Omron Sysmac Studio project 04820KA001 Mono Slitter 903_V12_1105 (Sysmac Studio 1.60.0.64010, StandardProject)
(* Modified to Connect 2nd Diameter Sens *)

# Controller PLC: NX1P2-9024DT1 version 1.42
Units and slaves: Node1 : IL EC BK-PAC(E001); 0 : IB IL 24 DI 8/HD-ECO(M1); 1 : IB IL 24 DO 8/HD-ECO(M2); Unit 1 : NX-PF0730 (N3); Unit 2 : NX-AD2603 (N1); Unit 3 : NX-EC0122 (N2)
Task PrimaryTask (priority 4, period or condition 4000): TaglMonoTRM

VAR_GLOBAL
    Pot1_Work_Velocity : INT;  (* Potentiometer 1 value - Work speed -	Valore potenziometro 1 - Lavoro -; at BuiltInIO://opt/#0/Ch1_Analog_Input_Value; published *)
    InvRef : INT;  (* Inverter speed reference	Riferimento velocità inverter; at BuiltInIO://opt/#0/Ch2_Analog_Output_Value; published *)
    Fix10Vdc : INT;  (* Fixed 10 Vdc generator	Generatore 10Vdc fisso; at BuiltInIO://opt/#0/Ch1_Analog_Output_Value; published *)
END_VAR
VAR_GLOBAL RETAIN
    VelMax : REAL := 800;  (* Maximum speed	Velocità massima; published *)
END_VAR
VAR_GLOBAL
    VelSet : REAL;  (* Set speed	Velocità impostata; published *)
END_VAR
VAR_GLOBAL RETAIN
    RwSlowDecelK : REAL := 0.15;  (* Learned slow-down decel per mm of rewinder diameter (mm/s2 per mm); published *)
    RwMaxSlowFallback : REAL := 1285.0;  (* Rewinder max: slow-down diameter while K not learned (mm); published *)
END_VAR
VAR_GLOBAL
    PaperDensity : REAL;  (* published *)
END_VAR
VAR_GLOBAL RETAIN
    Language : DINT;  (* Language	Lingua; published *)
    RwThickMin_mm : REAL := 0.02;  (* Learning: min plausible paper thickness (mm); published *)
END_VAR
VAR_GLOBAL
    PulseRate : UDINT;  (* Pulses per 100 ms	Impulsi * 100ms; at IOBus://unit#3/Ch1 Pulse Rate; published *)
END_VAR
VAR_GLOBAL RETAIN
    RwThickMax_mm : REAL := 2.0;  (* Learning: max plausible paper thickness (mm); published *)
    RwDecelMin_mm : REAL := 20.0;  (* Learning: min plausible stop decel (mm/s2); published *)
    RwDecelMax_mm : REAL := 5000.0;  (* Learning: max plausible stop decel (mm/s2); published *)
    RwLearnFailMax : INT := 12;  (* Learning: failed windows before alarm (12 = 2 min); published *)
    RwStopFailMax : INT := 3;  (* Learning: failed stops before alarm; published *)
    RwThick_mm : REAL;  (* Learned paper thickness (mm); published *)
END_VAR
VAR_GLOBAL
    OverSpeed : BOOL;  (* Speed too high	Velocità troppo alta; published *)
END_VAR
VAR_GLOBAL RETAIN
    WorkSpd_Max : REAL := 500.0;  (* Work speed pot full scale (m/min), 50..VelMax; published *)
    WorkSpd_Max_Set : REAL := 400.0;  (* HMI request: work pot full scale (m/min), applied only with motor stopped; published *)
    UwRawMin : INT := 10;  (* Unwinder sonar raw min (below = sensor fault, alarm 17); published *)
    UwRawMax : INT := 3990;  (* Unwinder sonar raw max (above = sensor fault / no echo, alarm 17); published *)
    TensCheckEnable : BOOL := False;  (* Tension check ON (HMI switch); OFF = start as before; published *)
    TensWaitSpd : REAL := 10.0;  (* Speed held after START until tension established (m/min); published *)
END_VAR
VAR_GLOBAL
    TensionOK : BOOL := False;  (* Tension established (debounced T-one Alarm 0); published *)
    TensWait : BOOL := False;  (* Waiting for tension (speed held at TensWaitSpd, HMI lamp); published *)
    SonarAsk : BOOL := False;  (* V10 HMI popup: sonar is OFF, turn it on? (HMI NO resets it); published *)
END_VAR
VAR_GLOBAL RETAIN
    UwSlow_at_D_Req : BOOL := True;  (* V7c: unwinder diameter slow-down follows the speed (FALSE = fixed UwSlowDown_Diam); published *)
END_VAR
VAR_GLOBAL
    UwSlowDiamAct : REAL := 0.0;  (* V7c: unwinder slows down at this diameter (mm), HMI display; published *)
END_VAR
VAR_GLOBAL RETAIN
    FinalStopDecel : REAL := 500.0;  (* V12: end-of-roll stop ramp, web decel (mm/s2), 0 = drive DEC ramp as before, 50..2000; published *)
END_VAR
VAR_GLOBAL
    FinalStopRamp : BOOL := False;  (* V12: end-of-roll stop ramp running (HMI lamp); published *)
END_VAR
VAR_GLOBAL RETAIN
    RwJogMaxDiam : REAL := 400.0;  (* V7d: jog blocked above this rewinder diameter (mm), 0 = no limit; published *)
END_VAR
VAR_GLOBAL
    JogInhibit : BOOL := False;  (* V7d: jog blocked (rewinder roll too big), HMI lamp; published *)
END_VAR
VAR_GLOBAL RETAIN
    SCurveTime : REAL := 0.5;  (* V7f: S-curve rounding of the AUTO ramps (s), 0 = off, max 2; published *)
END_VAR
VAR_GLOBAL
    TOneDecel : BOOL := False;  (* V7f: line decelerating (for a T-one stop/boost input); published *)
END_VAR
VAR_GLOBAL RETAIN
    HornStartBeep_s : REAL := 1.0;  (* V9 horn: beep when the slow-down starts (s), 0 = off, max 5; published *)
    HornBeepLen_s : REAL := 0.2;  (* V9 horn: length of the short beeps during slow-down (s), 0 = off, max 2; published *)
    HornBeepPeriod : REAL := 5.0;  (* V9 horn: one short beep every ... s during slow-down, 0 = off, max 30; published *)
    HornStopBeep_s : REAL := 3.0;  (* V9 horn: beep when stopped after a slow-down (s), 0 = off, max 10; published *)
END_VAR
VAR_GLOBAL
    HornTest : BOOL := False;  (* V9 horn: HMI test button (momentary), machine stopped only; published *)
END_VAR
VAR_GLOBAL RETAIN
    RwLockDiam : REAL := 300.0;  (* V9: paper thickness LOCKED at this rewinder diameter (mm), 0 = never lock; published *)
    RwLockMinGrow_mm : REAL := 50.0;  (* V9: min diameter growth since the start of learning before locking (mm); published *)
    RwMatLocked : BOOL := False;  (* V9: paper thickness locked (HMI lamp), NEW PAPER / GSM YES unlocks; published *)
END_VAR
VAR_GLOBAL
    LongThick_mm : REAL := 0.0;  (* V9: thickness from the long baseline (mm), HMI display; published *)
    RwDiamRev : REAL := 0.0;  (* V9: rewinder diameter averaged over one revolution (mm); published *)
    RwWave_mm : REAL := 0.0;  (* V9: diameter wave peak-peak in the last revolution (mm), HMI; published *)
    UwStopLenShow : BOOL := False;  (* V9 HMI: show unwinder STOP LENGTH (AUTO STOP UNWINDER active); published *)
    UwSlowDiamShow : BOOL := False;  (* V9 HMI: show unwinder SLOW AT diameter (normal operation, sonar ON); published *)
END_VAR
VAR_GLOBAL RETAIN
    SoftCancelAccel : REAL := 100.0;  (* V9: then ramp up at this web accel (mm/s2), 0 = AccelWeb; published *)
END_VAR
VAR_GLOBAL
    RwMatReset : BOOL := False;  (* HMI NEW PAPER: forget the learned paper thickness RwMat_K (PLC resets it); published *)
END_VAR
VAR_GLOBAL RETAIN
    FinalSpd_Max_Set : REAL := 80.0;  (* HMI request: final pot full scale (m/min), applied only with motor stopped; published *)
    FinalSpd_Max : REAL := 80.0;  (* Final speed pot full scale (m/min), 5..WorkSpd_Max; published *)
END_VAR
VAR_GLOBAL
    UnderSpeed : BOOL;  (* Speed too low	Velocità troppo bassa; published *)
    RwLearnReset : BOOL := False;  (* HMI / Watch: clear learned decels RwStopDecelK, RwStopDecel, RwSlowDecelK (PLC resets it); published *)
END_VAR
VAR_GLOBAL RETAIN
    RwCoreDiameter : REAL := 100.0;  (* Rewinder core outside diameter for TEACH CORE (mm); published *)
END_VAR
VAR_GLOBAL
    RwTeachCore : BOOL := False;  (* HMI: TEACH CORE request (PLC resets it); published *)
    RwTeachState : INT := 0;  (* TEACH CORE: 0 idle 1 teaching 2 done 3 refused; published *)
END_VAR
VAR_GLOBAL RETAIN
    SpdDelta_Percent : REAL := 12.0;  (* Speed difference percentage	Percentuale differenza velocità; published *)
END_VAR
VAR_GLOBAL
    Encoder_Pos : DINT;  (* Encoder counter	Contatore encoder; at IOBus://unit#3/Ch1 Encoder Present Position; published *)
    UwTeachState : INT := 0;  (* Unwinder TEACH CORE: 0 idle 1 teaching 2 done 3 refused; published *)
    Encoder_On : BOOL;  (* Encoder enable	Abilita encoder; at IOBus://unit#3/Ch1 Encoder Counter Operation Command/Ch1 Counter Enable; published *)
    Encoder_Reset : BOOL;  (* Encoder reset	Reset encoder; at IOBus://unit#3/Ch1 Encoder Counter Operation Command/Ch1 Internal Reset Execution; published *)
    HMI_Screen : ARRAY[0..1] OF DINT;  (* HMI panel Screen	Pagina pannello; published *)
END_VAR
VAR_GLOBAL RETAIN
    Velocity_M_min : REAL;  (* Speed in m/min	Velocità in mt/min; published *)
    Current_Metre : REAL;  (* Current metres	Metri attuali; published *)
END_VAR
VAR_GLOBAL
    I_RsetCnt : BOOL;  (* Metre counter reset button	Pulsante reset contametri; published *)
END_VAR
VAR_GLOBAL RETAIN
    Speed_Display : REAL;  (* Set speed (displayed)	Velocità impostata visualizzata; published *)
END_VAR
VAR_GLOBAL
    I_ControlVoltage : BOOL;  (* In_0 ControlVoltageON	Ausiliari inseriti; at BuiltInIO://cpu/#0/Input_Bit_00; published *)
    I_Start_PB : BOOL;  (* In_1 Start button	Pulsante di marcia; at BuiltInIO://cpu/#0/Input_Bit_01; published *)
    I_Stop_PB : BOOL;  (* In_2 Stop button	Pulsante di arresto; at BuiltInIO://cpu/#0/Input_Bit_02; published *)
    I_Motor_Thermal : BOOL;  (* In_3 Motor thermal switch	Pastiglia termica motore; at BuiltInIO://cpu/#0/Input_Bit_03; published *)
    I_Prot_ByPass : BOOL;  (* In_4 Guards-bypassed selector switch - Under Panel	Selettore protezioni escluse; at BuiltInIO://cpu/#0/Input_Bit_04; published *)
    I_Hub_Position : BOOL;  (* In_5 Hub/chuck in extraction position	Mozzo in posizione di estrazione; at BuiltInIO://cpu/#0/Input_Bit_05; published *)
    I_FrontGuard_Closed : BOOL;  (* In_6 Front guard closed	Riparo frontale chiuso; at BuiltInIO://cpu/#0/Input_Bit_06; published *)
    I_Jog_PB : BOOL;  (* In_7 Jog Push button	Pulsante velocità ridotta; at BuiltInIO://cpu/#0/Input_Bit_07; published *)
    I_VFD_Alarm : BOOL;  (* In_8 Inverter in alarm	Inverter in allarme; at BuiltInIO://cpu/#0/Input_Bit_08; published *)
    I_Side_Door_Closed : BOOL;  (* In_Side Door is Closed	Fotocellula diametro bobina; at BuiltInIO://cpu/#0/Input_Bit_13; published *)
    I_OR_Position_Sens : BOOL;  (* OverRider position sens	Sensore posizione pressore; at ECAT://node#[1,0]/IB IL 24 DI 8/HD-ECO Input-_IN01 (Pin 1.1)_6000_01; published *)
    I_OR_Hoover_Mode : BOOL;  (* OverRider Hoover Mode	Pressostato pressore; at ECAT://node#[1,0]/IB IL 24 DI 8/HD-ECO Input-_IN02 (Pin 2.1)_6000_02; published *)
    I_OR_Auto_OS : BOOL;  (* OverRider in automatic	Pressore in automatico; at ECAT://node#[1,0]/IB IL 24 DI 8/HD-ECO Input-_IN03 (Pin 1.2)_6000_03; published *)
    I_OR_Cont_OS : BOOL;  (* OverRider in continuous	Pressore in continuo; at ECAT://node#[1,0]/IB IL 24 DI 8/HD-ECO Input-_IN04 (Pin 2.2)_6000_04; published *)
    O_MotorStart : BOOL;  (* Q_0 Motor start	Start motore; at BuiltInIO://cpu/#0/Output_Bit_00; published *)
    I_FanTemp_Ok : BOOL;  (* Motor (fan) thermal OK	Termico motore ok; at ECAT://node#[1,0]/IB IL 24 DI 8/HD-ECO Input-_IN06 (Pin 2.3)_6000_06; published *)
    O_Alarm_Array : BOOL;  (* Alarm lamp	Lampada allarme; at ECAT://node#[1,1]/IB IL 24 DO 8/HD-ECO Output_OUT01 (Pin 1.1)_7000_01; published *)
    O_Prot_ByPass_Lamp : BOOL;  (* Guards bypassed lamp	Lampada protezioni escluse; published *)
    O_Motor_Lamp : BOOL;  (* Q_1 Motor ON lamp	Lampada motore on; at BuiltInIO://cpu/#0/Output_Bit_01; published *)
    O_RwUnload : BOOL;  (* Unloaders enable - opening	Consenso a scaricatori in apertura; at ECAT://node#[1,1]/IB IL 24 DO 8/HD-ECO Output_OUT03 (Pin 1.2)_7000_03; published *)
    O_FrontGuard_ByPass : BOOL;  (* Front guard bypass	Bypass protezione frontale; at ECAT://node#[1,1]/IB IL 24 DO 8/HD-ECO Output_OUT04 (Pin 2.2)_7000_04; published *)
    O_Brake : BOOL;  (* Q_2 Brake command	Comando freno; at BuiltInIO://cpu/#0/Output_Bit_02; published *)
    O_OR_Auto_Lamp : BOOL;  (* Q_6 OverRider auto/continuous lamp	Lamapda pressore in auto o continuo; at BuiltInIO://cpu/#0/Output_Bit_06; published *)
    O_OverRider_Up : BOOL;  (* Q_9 Raise OverRider ~10mm Over Rewinder roll	Solleva pressore; at BuiltInIO://cpu/#0/Output_Bit_09; published *)
    O_OverRider_Hold : BOOL;  (* Q_4 OverRider Lock 	Blocca pressore; at BuiltInIO://cpu/#0/Output_Bit_04; published *)
    O_CoolingFan : BOOL;  (* Q_3 Brake and motor fans	Ventole freno e motore; at BuiltInIO://cpu/#0/Output_Bit_03; published *)
END_VAR
VAR_GLOBAL RETAIN
    Fan_Timeout : REAL := 0.5;  (* Fans stop timeout [min]	Timeout stop ventole da pannello; published *)
    OverRider_TimeOFF : REAL := 0.01;  (* OverRider photocell OFF timeout (panel)	Timeout fotocellula pressore off; published *)
    OverRider_TimeON : REAL := 0.05;  (* OverRider photocell ON timeout (panel)	Timeout fotocellula pressore on; published *)
END_VAR
VAR_GLOBAL
    AlarmOn : BOOL;  (* Alarm active	Allarme presente; published *)
    BuzzerOn : BOOL;  (* Panel buzzer command	Comando buzzer pannello; published *)
    Msg : INT;  (* Message	Messagio; published *)
    Index_B : INT;  (* Alarm index	Indice allarme; published *)
    MotStop : BOOL;  (* Motor stopped	Motore fermo; published *)
    Clock1s : BOOL;  (* 1 s clock	Clock di 1s; published *)
END_VAR
VAR_GLOBAL RETAIN
    ManMode : BOOL;  (* Manual mode	Modo manuale; published *)
END_VAR
VAR_GLOBAL
    Counter_Reset : BOOL;  (* Counter reset from panel	Reset contatore da pannello; published *)
    I_FrontGuard_Open : BOOL;  (* In_9 Front guard open	Riparo frontale aperto; at BuiltInIO://cpu/#0/Input_Bit_09; published *)
    O_RwLoading_Enable : BOOL;  (* Q_7 Unloaders Load enable - closing	Consenso scaricatori in chiusura; at BuiltInIO://cpu/#0/Output_Bit_07; published *)
END_VAR
VAR_GLOBAL RETAIN
    JogSpd_SP : REAL := 10.0;  (* Speed in manual	Velocità in manuale; published *)
END_VAR
VAR_GLOBAL
    O_AccDec2 : BOOL;  (* Q_5 Second acc/dec ramp	Seconda rampa di acc/dec; at BuiltInIO://cpu/#0/Output_Bit_05; published *)
END_VAR
VAR_GLOBAL RETAIN
    AccelTrim : REAL := 0.08;  (* Acceleration coefficient in run	Coefficente accelerazione in lavoro; published *)
    DecelTrim : REAL := 0.08;  (* Deceleration coefficient in run	Coefficente decelerazione in lavoro; published *)
    DecelCoarse : REAL := 0.3;  (* Acceleration coefficient at start (orig. comment; name suggests decel)	Coefficente accelerazione in partenza; published *)
    AccelCoarse : REAL := 0.3;  (* Acceleration coefficient at start (orig. comment; name suggests accel)	Coefficente decelerazione in partenza; published *)
END_VAR
VAR_GLOBAL
    UwStopDiamShow : BOOL := False;  (* V11 HMI: show unwinder STOP AT diameter (slow-down reached, decel / final speed); published *)
    O_AcousticSignal : BOOL;  (* Q_8 Horn / Acoustic signal	Segnalatore acustico; at BuiltInIO://cpu/#0/Output_Bit_08; published *)
    Pot2_Slow_Velocity : INT;  (* Potentiometer 2 value - Final speed -	Valore potenziometro 2 - Finale -; at BuiltInIO://opt/#0/Ch2_Analog_Input_Value; published *)
    I_AutoStop_OS : BOOL;  (* In_10 Stop on metre counter	Arresto con contametri; at BuiltInIO://cpu/#0/Input_Bit_10; published *)
    I_Input_11_Spare_1255 : BOOL;  (* In_11 SPARE  (wire 12.55) Under Panel	Rallento a fine bobina; at BuiltInIO://cpu/#0/Input_Bit_11 *)
    I_WebBreak_Monitor : BOOL;  (* In_12 Paper break monitoring ON	Controllo rottura carta on; at BuiltInIO://cpu/#0/Input_Bit_12; published *)
    I_Vacuum_OK : BOOL;  (* Extractor fan thermal OK	Termico aspiratore ok; at IOBus://unit#3/Ch1 Reset/External Input Status/Ch1 External Input 0 Status; published *)
    I_T_one_TensionOK : BOOL;  (* T-one Alarm 0 (15-16): tension established (replaces I_SlowSens_PH); at ECAT://node#[1,0]/IB IL 24 DI 8/HD-ECO Input-_IN05 (Pin 1.3)_6000_05; published *)
    I_WebBreak_PH : BOOL;  (* Paper break photocell	Fotocellula rottura carta; at ECAT://node#[1,0]/IB IL 24 DI 8/HD-ECO Input-_IN07 (Pin 1.4)_6000_07; published *)
END_VAR
VAR_GLOBAL RETAIN
    UwStop_at_M_Val : REAL := 5100;  (* Unwinder Stop at metres	Metri totali; published *)
    UwSlowMargin_m : REAL := 10;  (* Unwinder Slow-down metres	Metri rallentamento; published *)
    LowSpd_Display : REAL;  (* Slow-down speed (displayed)	Velocità rallentamento visualizzata; published *)
    RwMaxDiam : REAL := 1315.0;  (* Rewinder max diameter protection (mm); published *)
END_VAR
VAR_GLOBAL
    RwMaxStop : BOOL;  (* Rewinder max diameter STOP (latched); published *)
END_VAR
VAR_GLOBAL RETAIN
    Encoder_Pulse : INT := 1000;  (* Encoder pulses/Rotation	Impulsi encoder; published *)
    RwSlowDecelLrn : REAL := 0.0;  (* Learned real slow-down decel (mm/s2) - 0 = not learned; published *)
END_VAR
VAR_GLOBAL
    CountReset_Req : BOOL;  (* Counter reset requested	Richiesto reset contatore; published *)
    Psw : INT;  (* Password Entry	Password; published *)
    I_RsetAlarm : BOOL;  (* Alarm reset	Reset allarmi; at ECAT://node#[1,0]/IB IL 24 DI 8/HD-ECO Input-_IN08 (Pin 2.4)_6000_08; published *)
END_VAR
VAR_GLOBAL RETAIN
    EncoderWheel_Circumf : REAL := 402;  (* Encoder wheel (Cylinder / Roller) Circumference [mm]	Diametro ruota encoder; published *)
END_VAR
VAR_GLOBAL
    AlarmCodeSV : ARRAY[0..32] OF BOOL;  (* Panel alarms	Allarmi a pannello; published *)
    SafeGuard_ByPass : BOOL;  (* Guards bypassed	Protezioni escluse; published *)
    FrontGuard_Closed : BOOL;  (* Front guard closed	Riparo frontale chiuso; published *)
    SoftStop : BOOL := False;  (* Soft stop in progress (HMI); published *)
END_VAR
VAR_GLOBAL RETAIN
    SoftStopEnable : BOOL := True;  (* STOP button = soft stop (False = immediate as before); published *)
    SoftStopEndSpd : REAL := 8.0;  (* Soft stop: run command drops below this speed (m/min); published *)
    UwDiam_Measure : REAL;  (* Measured distance	Distanza letta; published *)
    UwCoreDiameter : REAL := 100;  (* Core Outside diameter [mm]; published *)
    Core_Measure : BOOL := False;  (* Stored core value; published *)
    UwCoreDistance : REAL := 785.56;  (* Sonar distance to empty core. [mm]; published *)
END_VAR
VAR_GLOBAL
    AI_Diam_Unwinder : INT;  (* Analog value - UnWinder Diameter	Valore analogico misura bobina madre; at IOBus://unit#2/Ch1 Analog Input Value; published *)
END_VAR
VAR_GLOBAL RETAIN
    Measure_ON : BOOL := True;  (* Measurement enabled; published *)
    UwDiam_Act : REAL;  (* Measured roll diameter; published *)
    UwSlow_at_D_Val : REAL := 200;  (* Unwinder Slow-down diameter [mm]; published *)
    UwStopDiam_Limit : REAL := 110;  (* Stop diameter; published *)
END_VAR
VAR_GLOBAL
    Alarm_Reset : BOOL;  (* Alarm reset from panel; published *)
    Psw22 : BOOL;  (* Password 22 for Popup 22; published *)
    Psw44 : BOOL;  (* Password 44 for Popup 44; published *)
    I_Roll_OK : BOOL;  (* Roll OK / Broken Holder Joint; published *)
    AI_Diam_Rewinder : INT;  (* Analog value - ReWinder Diameter; at IOBus://unit#2/Ch2 Analog Input Value; published *)
END_VAR
VAR_GLOBAL RETAIN
    RwStopEnable : BOOL := False;  (* Rewinder diameter stop enabled; published *)
    RwTargetDiam : REAL := 300.0;  (* Rewinder final diameter (mm); published *)
    RwUseSlow : BOOL := True;  (* Slow down before target; published *)
    RwSlowMargin_m : REAL := 10.0;  (* Rewinder Metres at slow speed before stop; published *)
    RwSlowDecel : REAL := 0.0;  (* Rewinder Slow-down decel mm/s2 - 0 = auto from DecStart; published *)
    RwResetHyst : REAL := 50.0;  (* Reset requests below target - this [mm]; published *)
    RwDist0V : REAL := 0.0;  (* DT35 distance at 0 V (mm); published *)
    RwDist10V : REAL := 782.0;  (* DT35 distance at 10 V (mm); published *)
    RwRawMin : INT := 10;  (* Raw below = sensor fault; published *)
    RwRawMax : INT := 3900;  (* Raw above = sensor fault; published *)
END_VAR
VAR_GLOBAL
    RwStopOnFault : BOOL := True;  (* Stop on sensor fault; published *)
END_VAR
VAR_GLOBAL RETAIN
    RwAxisDist : REAL := 727.0;  (* Sensor to shaft centre (mm) - teach; published *)
    RwFilter_K : REAL := 0.2;  (* Distance filter per 100 ms (0..1); published *)
    RwMinPulses : DINT := 1000;  (* Min pulses in window to learn; published *)
    RwLearn_K : REAL := 0.3;  (* Material factor filter weight; published *)
    RwMat_K : REAL := 0.0;  (* Learned material factor; published *)
    RwLearnStop : BOOL := True;  (* Learn stop decel on every stop; published *)
    RwMinLearnSpd : REAL := 15.0;  (* Min speed to learn a stop (m/min); published *)
    RwStopDecel : REAL := 0.0;  (* Learned stop decel (pulses/s2); published *)
    RwTreact : REAL := 0.03;  (* Stop reaction time (s); published *)
    RwTstopDef : REAL := 3.0;  (* Stop time until decel learned (s); published *)
    RwTrim : REAL := 1.0;  (* Stop length trim (>1 = earlier); published *)
END_VAR
VAR_GLOBAL
    RwDist : REAL;  (* Filtered distance (mm); published *)
    RwDiam : REAL;  (* Rewinder diameter (mm); published *)
    RwSpeed : REAL;  (* Line speed from encoder (m/min); published *)
    RwRemain_m : REAL;  (* Metres to target diameter; published *)
    RwStopLen_m : REAL;  (* Stopping length now (m); published *)
    RwSlowLen_m : REAL;  (* Rewinder Slow-down length [m]; published *)
    RwStop_at_D_Req : BOOL;  (* Rewinder diameter STOP request; published *)
    RwSlow_at_D_Req : BOOL;  (* Rewinder diameter SLOW request; published *)
    RwSensFault : BOOL;  (* Rewinder DT35 sensor fault; published *)
END_VAR
VAR_GLOBAL RETAIN
    UwStopEnable : BOOL := False;  (* Unwinder Auto Stop - Enable; published *)
END_VAR
VAR_GLOBAL
    SlowAtDisp : REAL;  (* HMI: slow-down starts at (m or mm, see SlowAtMode); published *)
    SlowAtMode : INT;  (* HMI: 0=none 1=unwinder [m] 2=rewinder [mm]; published *)
    SlowAtShow : BOOL;  (* HMI: show slow-down display; published *)
    UwSlow_at_M_Val : REAL;  (* Unwinder: slow-down starts at [m]; published *)
    UwSlow_at_M_Req : BOOL;  (* Unwinder metre slow-down request (latched); published *)
    RwSlow_at_D_Val : REAL;  (* Rewinder slow-down starts at diameter [mm]; published *)
    RwStop_at_D_Val : REAL;  (* Rewinder: stop command at diameter (mm); published *)
    RwMaxSlow : BOOL;  (* Rewinder max diameter SLOW (latched); published *)
END_VAR
VAR_GLOBAL RETAIN
    UwEmptyHyst : REAL := 30.0;  (* Unwinder Empty Hysteresis; published *)
END_VAR
VAR_GLOBAL
    GSM_Learned_OK : BOOL;  (* Paper [Grams / Square Meter]  FALSE until GSM learned; published *)
    RwMaxSlowAtDiam : REAL := 1370.0;  (* Rewinder max: slow-down starts at diameter (mm); published *)
END_VAR
VAR_GLOBAL RETAIN
    RwStopDecelK : REAL := 0.0;  (* Learned stop decel per mm of rewinder diameter (mm/s2 per mm); published *)
    SoftStopDecel : REAL := 500.0;  (* Soft stop decel (mm/s2), 0 = DecelCoarse; published *)
END_VAR
VAR_GLOBAL
    SpdMax_Pending : BOOL := False;  (* New pot range waiting for the motor to stop; published *)
END_VAR
VAR_GLOBAL RETAIN
    RwAxisDist_Prev : REAL := 727.0;  (* Rewinder: RwAxisDist before the last TEACH (for UNDO); published *)
    UwCoreDist_Prev : REAL := 785.56;  (* Unwinder: UwCoreDistance before the last TEACH (for UNDO); published *)
END_VAR
VAR_GLOBAL
    RwTeachUndo : BOOL := False;  (* HMI: UNDO rewinder TEACH (PLC resets it); published *)
    UwTeachUndo : BOOL := False;  (* HMI: UNDO unwinder TEACH (PLC resets it); published *)
    Psw33 : BOOL;  (* Password 33 for Popup 33; published *)
END_VAR
VAR_GLOBAL RETAIN
    RwMatChangePct : REAL := 35.0;  (* Paper change detection: window deviation (%), 2 windows in a row = new paper, 0 = off; published *)
    RwSlowFallbackMm : REAL := 30.0;  (* Rewinder: slow-down this many mm before the target while the paper thickness is not learned (0 = off); published *)
    RwAutoMaxSpd : REAL := 500.0;  (* Rewinder AUTO stop ON: maximum work speed (m/min), 0 = no limit; published *)
    RwWinLen_m : REAL := 60.0;  (* Paper thickness learning: MAX window length (m of paper); published *)
    RwWinGrow_mm : REAL := 5;  (* Paper thickness learning: window = this diameter growth (mm), 4 m .. RwWinLen_m; published *)
END_VAR
VAR_GLOBAL
    GsmAsk : BOOL := False;  (* HMI popup: new parent roll, did you change the paper? (HMI NO resets it); published *)
    GsmAskYes : BOOL := False;  (* HMI popup YES: forget the learned thickness (PLC resets it); published *)
END_VAR
VAR_GLOBAL RETAIN
    DecelWeb : REAL := 250.0;  (* V7: AUTO decel ramp, real web mm/s2 (0 = DecelCoarse); published *)
    AccelWeb : REAL := 200.0;  (* AUTO accel ramp, real web mm/s2 (0 = AccelCoarse); published *)
    RwRatioD : REAL := 3366.0;  (* V7: drive counts per m/min x rewinder diameter (mm), adapted while running; published *)
    FFEnable : BOOL := True;  (* V7: feed-forward speed loop ON (FALSE = old loop of rung 16); published *)
END_VAR
VAR_GLOBAL
    SpdHold : BOOL := False;  (* V9: speed held after START during a soft stop, START again = ramp up (HMI lamp); published *)
    SonarAskYes : BOOL := False;  (* V10 HMI popup YES: sonar ON (PLC resets it); published *)
    UwStop_at_D_Val : REAL := 0.0;  (* V11: unwinder stop command diameter (mm) so the web stops at UwDiamStop, HMI "STOP AT"; published *)
    Clock10ms : BOOL;  (* 10mS clock; published *)
    Clock100ms : bool;  (* 100mS clock; published *)
    Sec_to_Min : REAL;
    Psw48 : BOOL;  (* Password 48 for Popup 48; published *)
    JogRun : BOOL;  (* V10: JOG really running (button, not a normal run, not a soft stop); published *)
    GuardStopOK : BOOL;  (* V11: stopped for real -> guard bypass allowed (Output 13); published *)
    SlowDown : BOOL;  (* Slow down	Rallenta; published *)
    WarningOn : bool;  (* HMI Warning Display; published *)
    AlarmSilenced : BOOL;  (* published *)
END_VAR
VAR_GLOBAL RETAIN
    PaperGSM : REAL;  (* published *)
    WebWidth_mm : REAL;  (* published *)
    TensFactor : REAL;  (* Tension Helper; published *)
    TensShowKg : BOOL;  (* Tension Helper; published *)
    TensShowLb : BOOL;  (* Tension Helper; published *)
    TensShowN : BOOL;  (* Tension Helper; published *)
    TensIdeal_Disp : REAL;  (* Tension Helper; published *)
    TensUnit : INT;  (* Tension Helper; published *)
END_VAR
VAR_GLOBAL
    TensUnitPB : BOOL;  (* Tension Helper; published *)
    TensLostWarn : BOOL := False;  (* Tension lost while running (warning); published *)
    UwSensTest : BOOL := False;  (* Unwinder sonar fault (raw out of range 1 s); published *)
    UwSensFault : BOOL;  (* UnWinder Sensor Fault; published *)
    Thickness_Fault : BOOL;  (* Thickness Not Learned !; published *)
    AutoStopWhy : INT;  (* published *)
    AutoStopDone : BOOL;  (* published *)
    AutoEnRefused : BOOL;  (* published *)
    AutoEnWhy : INT;  (* published *)
END_VAR

PROGRAM TaglMonoTRM
VAR
    SpdDelta : REAL;  (* Minimum or maximum speed SpdDeltaerence	Minima o massima differenza velocità *)
    UwSlowDiamCalc : REAL;  (* V7c: speed-dependent unwinder slow-down diameter (mm) *)
    SonarRunMem : bool;
    EndStopReq : BOOL;  (* V12: end-of-roll stop requested (AutoStopCmd or unwinder diameter) *)
    Buffer_R : BOOL;  (* Buffer Result *)
    EndRampOK : BOOL;  (* V12: end-of-roll ramp usable (FinalStopDecel, FF active, running) *)
    EndRampHard : BOOL;  (* V12: safety net during the ramp -> immediate stop *)
    EndStopNow : BOOL;  (* V12: immediate end-of-roll stop (Motor_Manager rung 4) *)
    SonarInit : bool;
    UwSlowDiamLatch : BOOL;  (* V7c: unwinder diameter slow-down reached (frozen) *)
    FFRate : REAL;  (* V7f: ramp rate (reference per 4 ms scan) *)
    FFRateSet : REAL;  (* V7f: rate allowed to still stop at the target *)
    FFJerk : REAL;  (* V7f: max rate change per scan *)
    SpdScanCnt : INT;  (* V9: scan counter for the 100 ms speed window *)
    HornRun : BOOL;  (* V9: slow-down / final speed running *)
    HornRunMem : BOOL;  (* V9: edge memory *)
    HornStartMem : BOOL;  (* V9: start edge memory *)
    HornTicks : INT;  (* V9: scans since slow-down start *)
    HornCnt : INT;  (* V9: scans in the beep period *)
    HornPer : INT;  (* V9: beep period in scans *)
    HornStartScans : INT;  (* V9: start beep in scans *)
    HornLenScans : INT;  (* V9: short beep in scans *)
    HornSlowBeep : BOOL;  (* V9: slow-down beep *)
    HornStopPend : BOOL;  (* V9: stopped after a slow-down, waiting for standstill *)
    HornStopTicks : INT;  (* V9: stop beep counter *)
    LongActive : BOOL;  (* V9: long-baseline learning running *)
    LongValid : BOOL;  (* V9: long baseline >= 20 mm growth, replaces the windows *)
    LongStartPos : DINT;  (* V9: encoder at the start of the long baseline *)
    LongStartD : REAL;  (* V9: rewinder diameter at the start (mm) *)
    LongGrow_mm : REAL;  (* V9: growth since the start (mm) *)
    LongPls : REAL;  (* V9: pulses since the start *)
    LongK : REAL;  (* V9: K from the long baseline *)
    RevW : REAL;  (* V9: encoder pulses summed in the current revolution *)
    RevDP : DINT;  (* V9: encoder pulses this scan *)
    RevPrevPos : DINT;  (* V9: encoder last scan *)
    RevSum : REAL;  (* V9: sum of raw DT35 distance x pulses *)
    RevMin : REAL;  (* V9: min raw distance in the revolution *)
    RevMax : REAL;  (* V9: max raw distance in the revolution *)
    RwDiamRevOk : BOOL;  (* V9: one full revolution averaged since the last fault *)
    UwEmptyTicks : INT;  (* V9: unwinder empty time (100 ms ticks) *)
    UwFullTicks : INT;  (* V9: new roll seen time (100 ms ticks) *)
    GsmArmed : BOOL;  (* V9: roll was empty -> next new roll asks the GSM question *)
    T_JogStartBlk : TOF;  (* V9: START blocked while JOG held + 2 s *)
    StartHeldBlk : BOOL;  (* V9: START pressed during the block, wait for release *)
    StartPB_OK : BOOL;  (* V9: START push-button accepted (replaces I_Start_PB in General 7/8/10) *)
    FFSoftMem : BOOL;  (* V9: soft stop last scan (rung B) *)
    FFSlowAcc : BOOL;  (* V9: gentle ramp-up after a cancelled soft stop *)
    FFStartEdge : BOOL;  (* V9: START push-button edge (rung B) *)
    FFStartMem : BOOL;  (* V9: START last scan (rung B) *)
    SpdDeltaMin : REAL;  (* Minimum speed difference	Minima differenza velocità *)
    FFSqrtArg : REAL;  (* SQRT argument (REAL) *)
    SpdDeltaMax : REAL;  (* Maximum speed SpdDeltaerence	Massima differenza velocità *)
    SoftStopMem : BOOL;  (* v6r: soft stop edge memory *)
    SoftStopRatio : REAL;  (* v6r: InvRef counts per m/min, frozen at the soft stop start *)
    MemPos : DINT;  (* Previous encoder count	Contatore encoder precedente *)
    MatChangeCnt : INT;  (* v6s: consecutive learning windows far from RwMat_K *)
    DeltaPulse : DINT;  (* Encoder count difference	Differenza contatore encoder *)
    SlowMem : BOOL;  (* SlowDown edge memory *)
    DecelDiam : REAL;  (* Rewinder diameter used by the decel model (mm, min 100) *)
    TeachSwap : REAL;  (* Temporary for UNDO swap *)
    SlowStartDiam : REAL;  (* Diameter at slow-down start (mm) *)
    BrakeHold : BOOL;  (* Keep T-one in auto during a normal stop (O_Brake) *)
    StopNow : BOOL;  (* Immediate stop request (replaces I_Stop_PB in General rung 9) *)
    StopPB_Mem : BOOL;  (* STOP button edge memory *)
    T_StopLong : TON;  (* STOP held 1 s = immediate stop *)
    T_SoftStop : TON;  (* Soft stop timeout (120 s) *)
    BrakeHoldTicks : INT;  (* BrakeHold duration after stop (100 ms ticks, max 150) *)
    StopStartDiam : REAL;  (* Diameter at stop command (mm) *)
    DecelK_Meas : REAL;  (* Measured decel per mm of diameter *)
    SlowMeasActive : BOOL;  (* Slow-down measurement running *)
    TeachTicks : INT;  (* TEACH CORE stable time (100 ms ticks) *)
    SlowStartPos : DINT;  (* Encoder at slow-down start *)
    SlowStartSpd_Pps : REAL;  (* Speed at slow-down start (pulses/s) *)
    SlowMeas_Pls : REAL;  (* Measured slow-down length (pulses) *)
    SlowDecelMeas_mm : REAL;  (* Measured slow-down decel (mm/s2) *)
    SlowOneRamp : BOOL;  (* Slow-down uses one ramp (manual or learned) *)
    Velocity : REAL;  (* Speed in [mm/s]	Velocità in mm/s *)
    Alarm_Array : ARRAY[0..32] OF BOOL;  (* Alarms	Allarme; [0] Not Used&#x9;pastiglia termica; [1] Motor fan thermal&#x9;termico ventola motore; [2] Inverter fault&#x9;anomalia inverter; [3] Emergency stop&#x9;in emergenza; [4] Motor thermal switch&#x9;pastiglia termica; [5] Front Guard moving&#x9;riparo in muovimento; [6] Web break&#x9;rottura carta; [7] Vacuum fan thermal&#x9;termico aspiratore; [8] Encoder Off&#x9;encoder fermo; [30] Hub not in position&#x9;Mozzo non in posizione; [9] Unloader Coupling Not Aligned; [10] Rewinder Diam Sensor Fault; [11] Rewinder max diam Protection.; [16] Rewinder GSM learning fault; [12] E-Stop by Holding Stop PB ; [13] Web Tension Too Low / Slack !; [14] UnWinder Diam Sensor Fault; [15] Unwinder Roll is Empty; [17] Thickness Not Learned !; [18] Side Door Opened; [19] Front Gate Not Closed !; [20] AutoStop Done !; [21] AutoStop Enable Monitor *)
    T_PlcOn : TON;  (* PLC active timeout	Timeout PLC attivo *)
    ControlVoltage : BOOL;  (* Auxiliaries OK	Ausiliari ok *)
    StartMotor_Cmd : BOOL;  (* Motor start command	Comando start motore *)
    HubExtractEnable : BOOL;  (* Hub extraction enable command	Comando consnso estrazione mozzo. *)
    Brake_Cmd : BOOL;  (* Brake command	Comando freno *)
    T_StopVent : TOF;  (* Fans stop timer	Timeout arresto ventole *)
    TimStopVen : TIME;  (* Fans stop timeout	Timeout stop ventole *)
    MotorCooling : BOOL;  (* Fans command	Comando ventole *)
    OverRider_Auto : BOOL;  (* OverRider in automatic	Pressore in automatico *)
    OverRider_Hoover : BOOL;  (* OverRider in Hoover Mode	Pressore in continuo *)
    OverRider_Lock : BOOL;  (* OverRider lock command	Comando blocco pressore *)
    GSM_LearnFault : BOOL;  (* Paper [Grams / Square Meter]   LearnFailCnt ≥ RwLearnFailMax *)
    TickCnt : INT;  (* 100 ms tick scan counter (25 x 4 ms) *)
    RunWasJog : BOOL;  (* Run used jog / manual / slow button (2nd ramp) *)
    StopLearnValid : BOOL;  (* This stop may be learned *)
    SpdBand_Pps : REAL;  (* Speed band of the trim ramp (pulses/s) *)
    TrimDecel_Pps2 : REAL;  (* Trim ramp decel (pulses/s2) *)
    SpdKnee_Pps : REAL;  (* Speed where coarse ramp hands over to trim ramp (pulses/s) *)
    OverRider_RaiseUp : BOOL;  (* OverRider raise command	Comando alzo pressore *)
    Pot1_Mem : INT;  (* Work potentiometer value	Valore potenziometro lavoro *)
    VelSet_mms : REAL;  (* Set speed in mm/s	Velocità impostata in mms *)
    Vfd_SP_Modif : REAL;  (* Inverter speed modifier	Modificatore velocità inverter *)
    RwAutoLimAct : BOOL;  (* v6y: rewinder AUTO speed limit active (taken over at standstill) *)
    UwTeachTicks : INT;  (* Unwinder TEACH CORE samples (100 ms) *)
    T_PosPresOff : TON;  (* OverRider photocell OFF timer	Timeout fotocellula pressore off *)
    T_PosPresOn : TON;  (* OverRider photocell ON timer	Timeout fotocellula pressore on *)
    TimPosPresOff : TIME;  (* OverRider photocell OFF timeout	Timeout fotocellula pressore off *)
    TimPosPresOn : TIME;  (* OverRider photocell ON timeout	Timeout fotocellula pressore on *)
    RollEnd_Active : BOOL;  (* Roll diameter photocell intercepted	Fotocellula diametro bobina intercettata *)
    Output_Ratio : REAL;  (* Analog output ratio	Rapporto analogica uscita *)
    Input_Ratio : REAL;  (* Analog input ratio	Rapporto analogica ingresso *)
    T_StartLow : TON;  (* Slow start timer	Timeout start lento *)
    T_UwDiamDebounce : TON;  (* Roll diameter photocell Debounce timer 500mS	Timeout fotocellula diamentro bobina off *)
    UwDiamReached : BOOL;  (* Roll diameter reached	Diamoetro bobina raggiunto *)
    Index_A : INT;
    AlarmStrobe : BOOL;  (* Alarm message display strobe	Strobe visualizza messagio allarme *)
    T_Display : TON;  (* Alarm display timer	Timeout visualizzazione allarme *)
    RangeOK : BOOL;  (* Range reached	Range raggiunto *)
    Vel_Max_mms : REAL;  (* Maximum speed in mm/s	Velocità massima in mm/sec *)
    Slow_Inhibit : BOOL;  (* Inhibit slow button	Inibisci pulsante slow *)
    Decel_Ramp : REAL;  (* Deceleration ramp	Rampa decelerazione *)
    Accel_Ramp : REAL;  (* Acceleration ramp	Rampa accelerazione *)
    Pot2_Mem : INT;  (* Final potentiometer value	Valore potenziometro finale *)
    Current_mm : REAL;  (* Current millimetres	Millimetri attuali *)
    EncoderPulse_to_mm : REAL;  (* mm per encoder pulse	mm per impulso encoder *)
    Stop : BOOL;  (* Stop	Arresto *)
    T_EncoderStill : TON;  (* (?) Encoder stopped timer *)
END_VAR
VAR RETAIN
    Analog_Res : UINT;  (* Analog board resolution	Risoluzione scheda analogica *)
END_VAR
VAR
    Mt_To_mm : REAL;  (* m/min to mm/s factor	Da Mt/min a mm/sec *)
END_VAR
VAR RETAIN
    Init_Ramp : BOOL;  (* (?) Ramp initialisation *)
END_VAR
VAR
    SlowByDiam : BOOL;  (* Slow down by diameter *)
    UwStopByDiam : BOOL;  (* Stop by diameter *)
    T_Screen_Delay : TON;  (* (?) Start page timer *)
    T_PulStop : TON;  (* (?) Stop button timer *)
END_VAR
VAR RETAIN
    Reading_Max : REAL := 2000;  (* Maximum sensor reading (full scale)	Lettura massima sensore *)
    DeadZone : REAL := 60;  (* Sensor dead zone	Zona morta sensore *)
    In_UwDiameter : REAL;  (* UnWinder Diameter Analog input voltage	Tensione ingresso analogico *)
END_VAR
VAR
    Tick : BOOL;  (* 100 ms tick *)
    MmPerPulse : REAL;  (* mm per encoder pulse *)
    RwDistRaw_mm : REAL;  (* Rewinder Unfiltered distance (mm) *)
    RwFiltInit : BOOL;  (* Rewinder Filter initialised *)
    SpdInit : BOOL;  (* Speed init *)
    EncPrev : DINT;  (* Encoder at previous tick *)
    SpdAct_Pps : REAL;  (* Actual Speed (pulses/s) *)
    LearnInit : BOOL;  (* Learn initialised *)
    LearnWinRunning : BOOL;  (* Motor ran whole window *)
    LearnWinTicks : INT;  (* Learn window counter *)
    LearnWin_Pls : DINT;  (* Pulses in window *)
    LearnWinDiamDelta : REAL;  (* Diameter change in window *)
    MatK_Window : REAL;  (* Material factor this window *)
    MotorRunMem : BOOL;  (* Motor start edge memory *)
    StopMeasActive : BOOL;  (* Stop measurement running *)
    StopStartPos : DINT;  (* Encoder at stop command *)
    StopStartSpd_Pps : REAL;  (* Speed at stop command (pulses/s) *)
    StandstillTicks : INT;  (* Standstill tick counter *)
    LearnWinOk : BOOL;  (* Learning window gave a valid result *)
    ThickWin_mm : REAL;  (* Paper thickness this window (mm) *)
    LearnFailCnt : INT;  (* Consecutive failed learning windows *)
    StopLearnOk : BOOL;  (* Stop measurement gave a valid result *)
    StopDecelMeas_mm : REAL;  (* Measured stop decel (mm/s2) *)
    StopMeas_Pls : REAL;  (* Measured stop length (pulses) *)
    StopDecelMeas : REAL;  (* Measured stop decel (pulses/s2) *)
    StopLen_Pls : REAL;  (* Stop length (pulses) *)
    StopLenFinal_Pls : REAL;  (* Stop length from slow speed (pulses) *)
    RwSlowLen_Pls : REAL;  (* Rewinder Slow-down length (pulses) *)
    SlowDecel_Pps2 : REAL;  (* Slow-down decel (pulses/s2) *)
    SpdFinal_Pps : REAL;  (* Final speed (pulses/s) *)
    RwRemain_Pls : REAL;  (* Rewinder Remaining length to target (pulses) *)
    LearnWinStartPos : DINT;  (* Rewinder Position Window 0 *)
    LearnWinStartDiam : REAL;  (* Rewinder Diameter Window 0 *)
    T_ByPassProtOff : TOF;  (* Delay Off Timer *)
    UwEnMem : BOOL;  (* Edge memory UwStopEnable *)
    RwEnMem : BOOL;  (* Edge memory RwEnable *)
    SpdRef_Pps : REAL;  (* Reference speed MAX(actual,setpoint) (pulses/s) *)
    SpdWork_Pps : REAL;  (* Work speed setpoint (pulses/s) *)
    SlowLenBase_Pls : REAL;  (* Slow-down length without margin (pulses) *)
    UwSlowLen_Pls : REAL;  (* Unwinder slow-down length (pulses) *)
    UwMarginUsed_m : REAL;  (* Unwinder margin at slow speed (m) *)
    SqrtArg : REAL;  (* Square root argument *)
    AutoSlowCmd : BOOL;  (* Automatic Slow Command *)
    AutoStopCmd : BOOL;  (* Automatic Stop Command *)
    RwLastValidDiam : REAL;  (* Rewinder Last valid diameter (mm) *)
    RwRemainMax_Pls : REAL;  (* Rewinder Remaining length to max diameter (pulses) *)
    UnWinder_Empty : BOOL;  (* UnWinder Empty *)
    StopFailCnt : INT;  (* Consecutive failed stop measurements *)
    UwTeachSum : REAL;  (* Unwinder TEACH CORE sonar sum (mm) *)
    T_MatReset : TON;  (* v6s: RwMatReset stays ON 3 s *)
    RwAutoMaxSpdAct : REAL;  (* v6y: active rewinder AUTO max speed (taken over at standstill) *)
    UwEmptyMem : BOOL;  (* v6x: UnWinder_Empty edge memory *)
    LearnWinLen_Pls : REAL;  (* v6w: learning window length in encoder pulses *)
    WebRatio : REAL;  (* V7: drive counts per m/min of web at the current diameter *)
    FFActive : BOOL;  (* V7: feed-forward loop active *)
    FFWasActive : BOOL;  (* V7: edge memory *)
    FFTarget : REAL;  (* V7: reference for the set speed (mm/s of the 0-10 V scale) *)
    RampRef : REAL;  (* V7: ramped reference (mm/s of the 0-10 V scale) *)
    StepAcc : REAL;  (* V7: accel step per scan *)
    StepDec : REAL;  (* V7: decel step per scan *)
    FFSteadyTicks : INT;  (* V7: scans at target *)
    FFErr : REAL;  (* V7: relative speed error *)
    Clock_100ms : bool;  (* Clock100ms *)
    AlarmCnt : INT;
    AlarmCntMem : INT;
    RstEdge : BOOL;
    RstMem : BOOL;
    SilenceTicks : INT;
    WarnCnt : INT;
    WarnCntMem : INT;
    WarnBeepTicks : INT;
    TensUnitMem : BOOL;
    TensIdeal_N : REAL;
    TensionSeen : BOOL := False;  (* Tension reached once since START *)
    T_TensOn : TON;  (* Tension ON debounce 0.5 s *)
    T_TensOff : TON;  (* Tension OFF debounce 2 s *)
    T_UwSensFlt : TON;  (* Unwinder sonar fault debounce 1 s *)
    Buffer_A : BOOL;
    Buffer_B : BOOL;
    Buffer_C : BOOL;
    Buffer_D : BOOL;
    AS_RunMem : BOOL;
    AutoStopSeen : BOOL;
    T_AutoStopDisp : TON;
    RwArmMem : BOOL;
    UwArmMem : BOOL;
    T_AutoEnRef : TON;
END_VAR
VAR_EXTERNAL
    VelSet : REAL;  (* Set speed *)
    OverSpeed : BOOL;  (* Speed too high *)
    SpdDelta_Percent : REAL;  (* Speed difference percentage *)
    Encoder_Pos : DINT;  (* Encoder counter *)
    FinalStopDecel : REAL;
    FinalStopRamp : BOOL;
    Velocity_M_min : REAL;  (* Speed in m/min *)
    Current_Metre : REAL;  (* Current metres	Metri attuali *)
    I_RsetCnt : BOOL;  (* Metre counter reset button *)
    SonarAsk : BOOL;
    SonarAskYes : BOOL;
    WorkSpd_Max_Set : REAL;  (* HMI request: work pot full scale (m/min), applied only with motor stopped *)
    FinalSpd_Max_Set : REAL;  (* HMI request: final pot full scale (m/min), applied only with motor stopped *)
    SpdMax_Pending : BOOL;  (* New pot range waiting for the motor to stop *)
    RwAxisDist_Prev : REAL;  (* Rewinder: RwAxisDist before the last TEACH (for UNDO) *)
    UwCoreDist_Prev : REAL;  (* Unwinder: UwCoreDistance before the last TEACH (for UNDO) *)
    RwTeachUndo : BOOL;  (* HMI: UNDO rewinder TEACH (PLC resets it) *)
    UwTeachUndo : BOOL;  (* HMI: UNDO unwinder TEACH (PLC resets it) *)
    RwLearnReset : BOOL;  (* HMI / Watch: clear learned decels RwStopDecelK, RwStopDecel, RwSlowDecelK (PLC resets it) *)
    UnderSpeed : BOOL;  (* Speed too low *)
    I_ControlVoltage : BOOL;  (* Auxiliaries ON *)
    I_Side_Door_Closed : BOOL;  (* Roll diameter photocell *)
    RwCoreDiameter : REAL;  (* Rewinder core outside diameter for TEACH CORE (mm) *)
    UwTeachState : INT;  (* Unwinder TEACH CORE: 0 idle 1 teaching 2 done 3 refused *)
    SoftStop : BOOL;  (* Soft stop in progress (HMI) *)
    SoftStopEnable : BOOL;  (* STOP button = soft stop (False = immediate as before) *)
    SoftStopEndSpd : REAL;  (* Soft stop: run command drops below this speed (m/min) *)
    SoftStopDecel : REAL;  (* Soft stop decel (mm/s2), 0 = DecelCoarse *)
    RwTeachCore : BOOL;  (* HMI: TEACH CORE request (PLC resets it) *)
    RwTeachState : INT;  (* TEACH CORE: 0 idle 1 teaching 2 done 3 refused *)
    O_MotorStart : BOOL;  (* Motor start *)
    RwSlowDecelK : REAL;  (* Learned slow-down decel per mm of rewinder diameter (mm/s2 per mm) *)
    RwStopDecelK : REAL;  (* Learned stop decel per mm of rewinder diameter (mm/s2 per mm) *)
    I_OR_Position_Sens : BOOL;  (* Rider roll position sensor *)
    WorkSpd_Max : REAL;  (* Work speed pot full scale (m/min), 50..VelMax *)
    FinalSpd_Max : REAL;  (* Final speed pot full scale (m/min), 5..WorkSpd_Max *)
    I_OR_Hoover_Mode : BOOL;  (* Rider roll pressure switch *)
    I_OR_Auto_OS : BOOL;  (* Rider roll in automatic *)
    I_OR_Cont_OS : BOOL;  (* Rider roll in continuous *)
    I_Start_PB : BOOL;  (* Start button *)
    I_Motor_Thermal : BOOL;  (* Motor thermal switch *)
    I_FanTemp_Ok : BOOL;  (* Motor (fan) thermal OK *)
    I_Stop_PB : BOOL;  (* Stop button *)
    I_Hub_Position : BOOL;  (* Hub/chuck in extraction position *)
    I_FrontGuard_Closed : BOOL;  (* Front guard closed *)
    RwMaxSlowFallback : REAL;  (* Rewinder max: slow-down diameter while K not learned (mm) *)
    RwMaxSlowAtDiam : REAL;  (* Rewinder max: slow-down starts at diameter (mm) *)
    O_Alarm_Array : BOOL;  (* Alarm lamp *)
    O_RwUnload : BOOL;  (* Unloaders enable - opening *)
    I_Prot_ByPass : BOOL;  (* Guards-bypassed selector switch *)
    O_Prot_ByPass_Lamp : BOOL;  (* Guards bypassed lamp *)
    O_Brake : BOOL;  (* Brake command *)
    Fan_Timeout : REAL;  (* Fans stop timeout (from panel) *)
    O_CoolingFan : BOOL;  (* Brake and motor fans *)
    O_OR_Auto_Lamp : BOOL;  (* Rider roll auto/continuous lamp *)
    O_OverRider_Up : BOOL;  (* Raise rider roll *)
    O_OverRider_Hold : BOOL;  (* Lock rider roll *)
    Fix10Vdc : INT;  (* Fixed 10 Vdc generator *)
    InvRef : INT;  (* Inverter speed reference *)
    Encoder_On : BOOL;  (* Encoder enable *)
    Encoder_Reset : BOOL;  (* Encoder reset *)
    OverRider_TimeOFF : REAL;  (* Rider roll photocell OFF timeout (panel) *)
    OverRider_TimeON : REAL;  (* Rider roll photocell ON timeout (panel) *)
    VelMax : REAL;  (* Maximum speed *)
    I_Jog_PB : BOOL;  (* Slow speed button *)
    O_Motor_Lamp : BOOL;  (* Motor ON lamp *)
    AlarmOn : BOOL;  (* Alarm active	Allarme presente *)
    BuzzerOn : BOOL;  (* Panel buzzer command	Comando buzzer pannelli *)
    I_VFD_Alarm : BOOL;  (* Inverter in alarm *)
    Msg : INT;  (* Message	Messaggio *)
    Index_B : INT;  (* Active alarm index	Indice allarme presente *)
    MotStop : BOOL;  (* Motor stopped	Motore in stop *)
    Clock1s : BOOL;  (* 1 s clock	Clock di 1s *)
    ManMode : BOOL;  (* Manual mode	Modo manuale *)
    Counter_Reset : BOOL;  (* Panel counter reset button	Pulsante reset contatore pannello *)
    I_FrontGuard_Open : BOOL;  (* Front guard open *)
    O_RwLoading_Enable : BOOL;  (* Unloaders enable - closing *)
    JogSpd_SP : REAL;  (* Speed in manual *)
    O_AccDec2 : BOOL;  (* Second acc/dec ramp *)
    AccelTrim : REAL;  (* Acceleration coefficient in run *)
    DecelTrim : REAL;  (* Deceleration coefficient in run *)
    DecelCoarse : REAL;  (* Acceleration coefficient at start (orig. comment; name suggests decel) *)
    AccelCoarse : REAL;  (* Deceleration coefficient at start (orig. comment; name suggests accel) *)
    Speed_Display : REAL;  (* Set speed (displayed) *)
    O_AcousticSignal : BOOL;  (* Horn / acoustic signal *)
    Pot1_Work_Velocity : INT;  (* Potentiometer 1 value - Work speed - *)
    O_FrontGuard_ByPass : BOOL;  (* Front guard bypass *)
    Pot2_Slow_Velocity : INT;  (* Potentiometer 2 value - Final speed - *)
    LowSpd_Display : REAL;  (* Slow-down speed (displayed) *)
    Encoder_Pulse : INT;  (* Encoder pulses *)
    RwSlowDecelLrn : REAL;  (* Learned real slow-down decel (mm/s2) - 0 = not learned *)
    UwSlowMargin_m : REAL;  (* Slow-down metres *)
    UwStop_at_M_Val : REAL;  (* Total metres *)
    I_AutoStop_OS : BOOL;  (* Stop on metre counter *)
    I_Input_11_Spare_1255 : BOOL;  (* Slow down at end of roll *)
    I_T_one_TensionOK : BOOL;  (* Slow-down photocell *)
    I_WebBreak_Monitor : BOOL;  (* Paper break monitoring ON *)
    I_WebBreak_PH : BOOL;  (* Paper break photocell *)
    I_Vacuum_OK : BOOL;  (* Extractor fan thermal OK *)
    CountReset_Req : BOOL;  (* Metre counter reset request	Richiesta azzeramento contametri *)
    Psw : INT;  (* Password *)
    I_RsetAlarm : BOOL;  (* Alarm reset *)
    EncoderWheel_Circumf : REAL;  (* Encoder wheel diameter *)
    AlarmCodeSV : ARRAY[0..32] OF BOOL;  (* Panel alarms *)
    SafeGuard_ByPass : BOOL;  (* Guards bypassed *)
    FrontGuard_Closed : BOOL;  (* Front guard closed *)
    Core_Measure : BOOL;  (* (?) Stored core value *)
    UwDiam_Measure : REAL;  (* Measured distance *)
    UwCoreDistance : REAL;  (* (?) Core measurement *)
    RwSlowFallbackMm : REAL;
    AI_Diam_Unwinder : INT;  (* Analog value - parent roll measurement *)
    RwMatChangePct : REAL;
    UwCoreDiameter : REAL;  (* (?) Shaft diameter *)
    Measure_ON : BOOL;  (* (?) Measurement enabled *)
    UwDiam_Act : REAL;  (* (?) Measured roll diameter *)
    UwStopDiam_Limit : REAL;  (* (?) Stop diameter *)
    UwSlow_at_D_Val : REAL;  (* (?) Slow-down diameter *)
    Alarm_Reset : BOOL;  (* (?) Alarm reset from panel *)
    HMI_Screen : ARRAY[0..1] OF DINT;  (* HMI panel page *)
    Psw22 : BOOL;  (* (?) Password 22 *)
    RwMatReset : BOOL;
    Psw44 : BOOL;  (* (?) Password 44 *)
    I_Roll_OK : BOOL;  (* (?) Roll OK *)
    AI_Diam_Rewinder : INT;  (* Rewinder DT35 raw - I/O Map Unit2 Ch2 *)
    RwStopEnable : BOOL;  (* Rewinder diameter stop enabled *)
    RwTargetDiam : REAL;  (* Rewinder final diameter (mm) *)
    RwUseSlow : BOOL;  (* Slow down before target *)
    RwSlowMargin_m : REAL;  (* Metres at slow speed before stop *)
    UwRawMin : INT;
    UwRawMax : INT;
    RwSlowDecel : REAL;  (* Slow-down decel mm/s2 - 0 = auto from DecStart *)
    RwResetHyst : REAL;  (* Reset requests below target - this (mm) *)
    RwDist0V : REAL;  (* DT35 distance at 0 V (mm) *)
    RwDist10V : REAL;  (* DT35 distance at 10 V (mm) *)
    RwRawMin : INT;  (* Raw below = sensor fault *)
    RwRawMax : INT;  (* Raw above = sensor fault *)
    RwStopOnFault : BOOL;  (* Stop on sensor fault *)
    RwAxisDist : REAL;  (* Sensor to shaft centre (mm) - teach *)
    RwFilter_K : REAL;  (* Distance filter per 100 ms (0..1) *)
    RwMinPulses : DINT;  (* Min pulses in window to learn *)
    RwLearn_K : REAL;  (* Material factor filter weight *)
    RwMat_K : REAL;  (* Learned material factor *)
    RwLearnStop : BOOL;  (* Learn stop decel on every stop *)
    RwMinLearnSpd : REAL;  (* Min speed to learn a stop (m/min) *)
    RwStopDecel : REAL;  (* Learned stop decel (pulses/s2) *)
    RwTreact : REAL;  (* Stop reaction time (s) *)
    RwTstopDef : REAL;  (* Stop time until decel learned (s) *)
    RwTrim : REAL;  (* Stop length trim (>1 = earlier) *)
    RwDist : REAL;  (* Filtered distance (mm) *)
    RwDiam : REAL;  (* Rewinder diameter (mm) *)
    RwSpeed : REAL;  (* Line speed from encoder (m/min) *)
    RwRemain_m : REAL;  (* Metres to target diameter *)
    RwStopLen_m : REAL;  (* Stopping length now (m) *)
    RwSlowLen_m : REAL;  (* Slow-down length now (m) *)
    RwStop_at_D_Req : BOOL;  (* Rewinder diameter STOP request *)
    RwSlow_at_D_Req : BOOL;  (* Rewinder diameter SLOW request *)
    RwSensFault : BOOL;  (* Rewinder DT35 sensor fault *)
    UwStopEnable : BOOL;  (* Unwinder metre-counter stop ON (HMI) *)
    SlowAtDisp : REAL;  (* HMI: slow-down starts at (m or mm, see SlowAtMode) *)
    UwSlow_at_D_Req : BOOL;
    UwSlowDiamAct : REAL;
    RwJogMaxDiam : REAL;
    JogInhibit : BOOL;
    SCurveTime : REAL;
    TOneDecel : BOOL;
    HornStartBeep_s : REAL;
    HornBeepLen_s : REAL;
    HornBeepPeriod : REAL;
    HornStopBeep_s : REAL;
    HornTest : BOOL;
    RwLockDiam : REAL;
    UwSensTest : BOOL;
    RwLockMinGrow_mm : REAL;
    RwMatLocked : BOOL;
    LongThick_mm : REAL;
    RwDiamRev : REAL;
    RwWave_mm : REAL;
    UwStopLenShow : BOOL;
    UwSlowDiamShow : BOOL;
    SoftCancelAccel : REAL;
    SpdHold : BOOL;
    SlowAtMode : INT;  (* HMI: 0=none 1=unwinder [m] 2=rewinder [mm] *)
    SlowAtShow : BOOL;  (* HMI: show slow-down display *)
    UwSlow_at_M_Val : REAL;  (* Unwinder: slow-down starts at (m) *)
    UwSlow_at_M_Req : BOOL;  (* Unwinder metre slow-down request (latched) *)
    RwSlow_at_D_Val : REAL;  (* Rewinder: slow-down starts at diameter (mm) *)
    RwStop_at_D_Val : REAL;  (* Rewinder: stop command at diameter (mm) *)
    RwMaxDiam : REAL;  (* Rewinder max diameter protection (mm) *)
    RwMaxStop : BOOL;  (* Rewinder max diameter STOP (latched) *)
    RwMaxSlow : BOOL;  (* Rewinder max diameter SLOW (latched) *)
    UwEmptyHyst : REAL;
    RwThickMin_mm : REAL;  (* Learning: min plausible paper thickness (mm) *)
    RwThickMax_mm : REAL;  (* Learning: max plausible paper thickness (mm) *)
    RwDecelMin_mm : REAL;  (* Learning: min plausible stop decel (mm/s2) *)
    RwDecelMax_mm : REAL;  (* Learning: max plausible stop decel (mm/s2) *)
    RwLearnFailMax : INT;  (* Learning: failed windows before alarm (12 = 2 min) *)
    RwStopFailMax : INT;  (* Learning: failed stops before alarm *)
    GSM_Learned_OK : BOOL;  (* Rewinder learning fault (alarm 16) *)
    RwThick_mm : REAL;  (* Learned paper thickness (mm) *)
    Psw33 : BOOL;
    RwAutoMaxSpd : REAL;
    RwWinLen_m : REAL;
    RwWinGrow_mm : REAL;
    GsmAsk : BOOL;
    GsmAskYes : BOOL;
    DecelWeb : REAL;
    AccelWeb : REAL;
    RwRatioD : REAL;
    FFEnable : BOOL;
    UwStopDiamShow : BOOL;
    UwStop_at_D_Val : REAL;
    Clock10ms : BOOL;
    Sec_to_Min : REAL;
    Psw48 : BOOL;
    JogRun : BOOL;
    GuardStopOK : BOOL;  (* V11: stopped for real -> guard bypass allowed (Output 13) *)
    SlowDown : BOOL;  (* Slow down	Rallenta *)
    WarningOn : bool;
    AlarmSilenced : BOOL;
    PaperGSM : REAL;
    WebWidth_mm : REAL;
    TensFactor : REAL;
    TensShowKg : BOOL;
    TensShowLb : BOOL;
    TensShowN : BOOL;
    TensIdeal_Disp : REAL;
    TensUnit : INT;
    TensUnitPB : BOOL;
    TensCheckEnable : BOOL;
    TensLostWarn : BOOL;
    TensWaitSpd : REAL;
    TensWait : BOOL;
    TensionOK : BOOL;
    UwSensFault : BOOL;
    Thickness_Fault : BOOL;
    AutoStopDone : BOOL;
    AutoStopWhy : INT;
    AutoEnRefused : BOOL;
    AutoEnWhy : INT;
END_VAR
VAR
    _p1 : BOOL;
    _e2 : R_TRIG;
    _e3 : F_TRIG;
    _p4 : BOOL;
    _p5 : BOOL;
    _p6 : BOOL;
    _p7 : BOOL;
    _e8 : R_TRIG;
    _e9 : R_TRIG;
    _e10 : R_TRIG;
    _e11 : R_TRIG;
    _e12 : R_TRIG;
    _e13 : R_TRIG;
    _e14 : F_TRIG;
END_VAR

(* Section General: ladder, written here as Structured Text *)

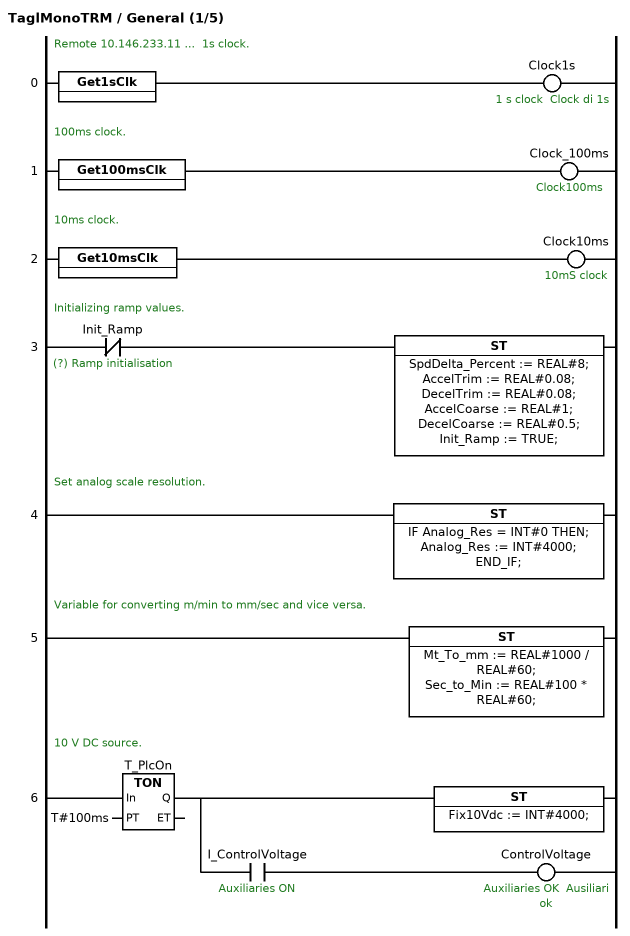
(* Rung 0: Remote 10.146.233.11 ...  1s clock. *)
Clock1s := Get1sClk();
(* Rung 1: 100ms clock. *)
Clock_100ms := Get100msClk();
(* Rung 2: 10ms clock. *)
Clock10ms := Get10msClk();
(* Rung 3: Initializing ramp values. *)
_p1 := NOT Init_Ramp;
IF _p1 THEN
    SpdDelta_Percent := REAL#8;
    AccelTrim := REAL#0.08;
    DecelTrim := REAL#0.08;
    AccelCoarse := REAL#1;
    DecelCoarse := REAL#0.5;
    Init_Ramp := TRUE;
END_IF;
(* Rung 4: Set analog scale resolution. *)
IF Analog_Res = INT#0 THEN;
	Analog_Res := INT#4000;
END_IF;
(* Rung 5: Variable for converting m/min to mm/sec and vice versa. *)
Mt_To_mm := REAL#1000 / REAL#60;
Sec_to_Min := REAL#100 * REAL#60;
(* Rung 6: 10 V DC source. *)
T_PlcOn(In := TRUE, PT := T#100ms);
IF T_PlcOn.Q THEN
    Fix10Vdc := INT#4000;
END_IF;
ControlVoltage := T_PlcOn.Q AND I_ControlVoltage;

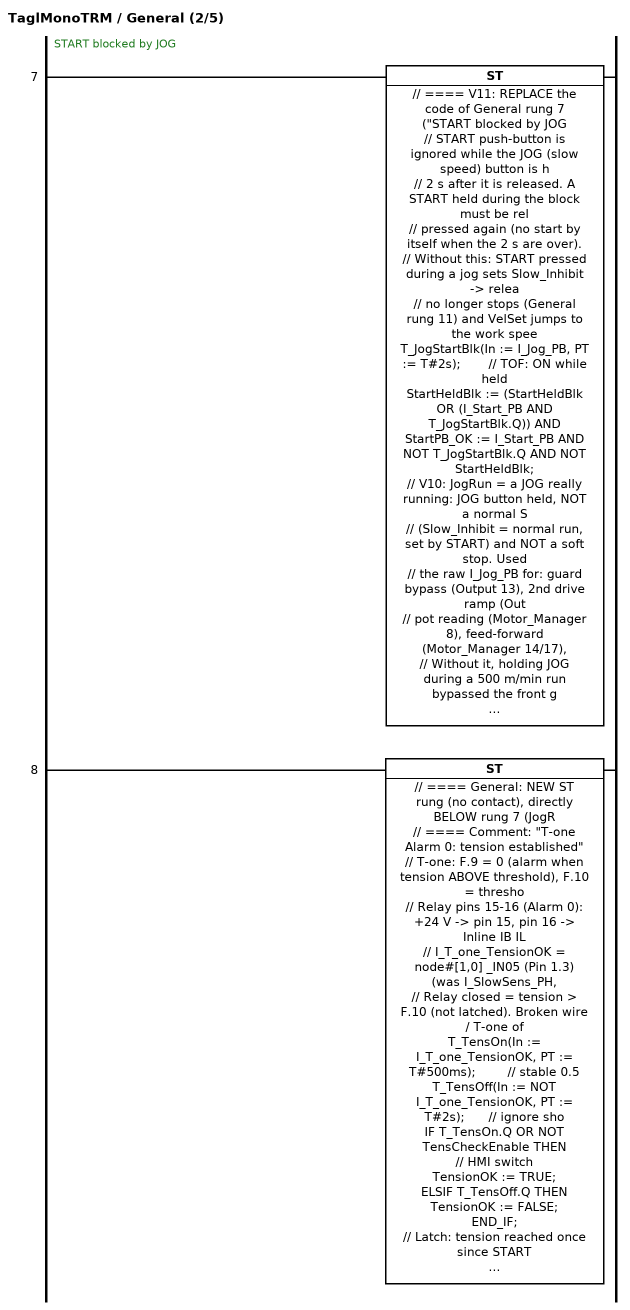
(* Rung 7: START blocked by JOG *)
// ==== V11: REPLACE the code of General rung 7 ("START blocked by JOG", printed V9).
// START push-button is ignored while the JOG (slow speed) button is held and for
// 2 s after it is released. A START held during the block must be released and
// pressed again (no start by itself when the 2 s are over).
// Without this: START pressed during a jog sets Slow_Inhibit -> releasing the jog
// no longer stops (General rung 11) and VelSet jumps to the work speed.

T_JogStartBlk(In := I_Jog_PB, PT := T#2s);       // TOF: ON while held + 2 s
StartHeldBlk := (StartHeldBlk OR (I_Start_PB AND T_JogStartBlk.Q)) AND I_Start_PB;
StartPB_OK := I_Start_PB AND NOT T_JogStartBlk.Q AND NOT StartHeldBlk;

// V10: JogRun = a JOG really running: JOG button held, NOT a normal START run
// (Slow_Inhibit = normal run, set by START) and NOT a soft stop. Used instead of
// the raw I_Jog_PB for: guard bypass (Output 13), 2nd drive ramp (Output 12),
// pot reading (Motor_Manager 8), feed-forward (Motor_Manager 14/17), AutoStop learning.
// Without it, holding JOG during a 500 m/min run bypassed the front gate / lateral
// doors safety (23KA4 // 5SA1) and switched the drive to its 2nd ramp.

JogRun := I_Jog_PB AND NOT Slow_Inhibit AND NOT SoftStop;

// Guard bypass (Output_Manager rung 13, 23KA4 // 5SA1): ON when the run command is
// off (machine stopped by the operator).

GuardStopOK := NOT StartMotor_Cmd;
(* Rung 8 *)
// ==== General: NEW ST rung (no contact), directly BELOW rung 7 (JogRun / GuardStopOK)
// ==== Comment: "T-one Alarm 0: tension established"
// T-one: F.9 = 0 (alarm when tension ABOVE threshold), F.10 = threshold (kg), F.11 = full scale
// Relay pins 15-16 (Alarm 0): +24 V -> pin 15, pin 16 -> Inline IB IL 24 DI 8 IN05, pin 1.3
// I_T_one_TensionOK = node#[1,0] _IN05 (Pin 1.3) (was I_SlowSens_PH, used in no rung)
// Relay closed = tension > F.10 (not latched). Broken wire / T-one off = "no tension" (fail-safe).

T_TensOn(In := I_T_one_TensionOK, PT := T#500ms);        // stable 0.5 s
T_TensOff(In := NOT I_T_one_TensionOK, PT := T#2s);      // ignore short dips (splice, wave, chatter)

IF T_TensOn.Q OR NOT TensCheckEnable THEN                // HMI switch OFF = old behaviour
    TensionOK := TRUE;
ELSIF T_TensOff.Q THEN
    TensionOK := FALSE;
END_IF;

// Latch: tension reached once since START

IF NOT StartMotor_Cmd THEN
    TensionSeen := FALSE;
ELSIF TensionOK THEN
    TensionSeen := TRUE;
END_IF;

// After START: hold at TensWaitSpd until the tension is there (JOG not affected)

TensWait := StartMotor_Cmd AND NOT TensionSeen AND NOT JogRun;

// Tension lost later while running -> warning only (no slow-down)

TensLostWarn := StartMotor_Cmd AND TensionSeen AND NOT TensionOK;

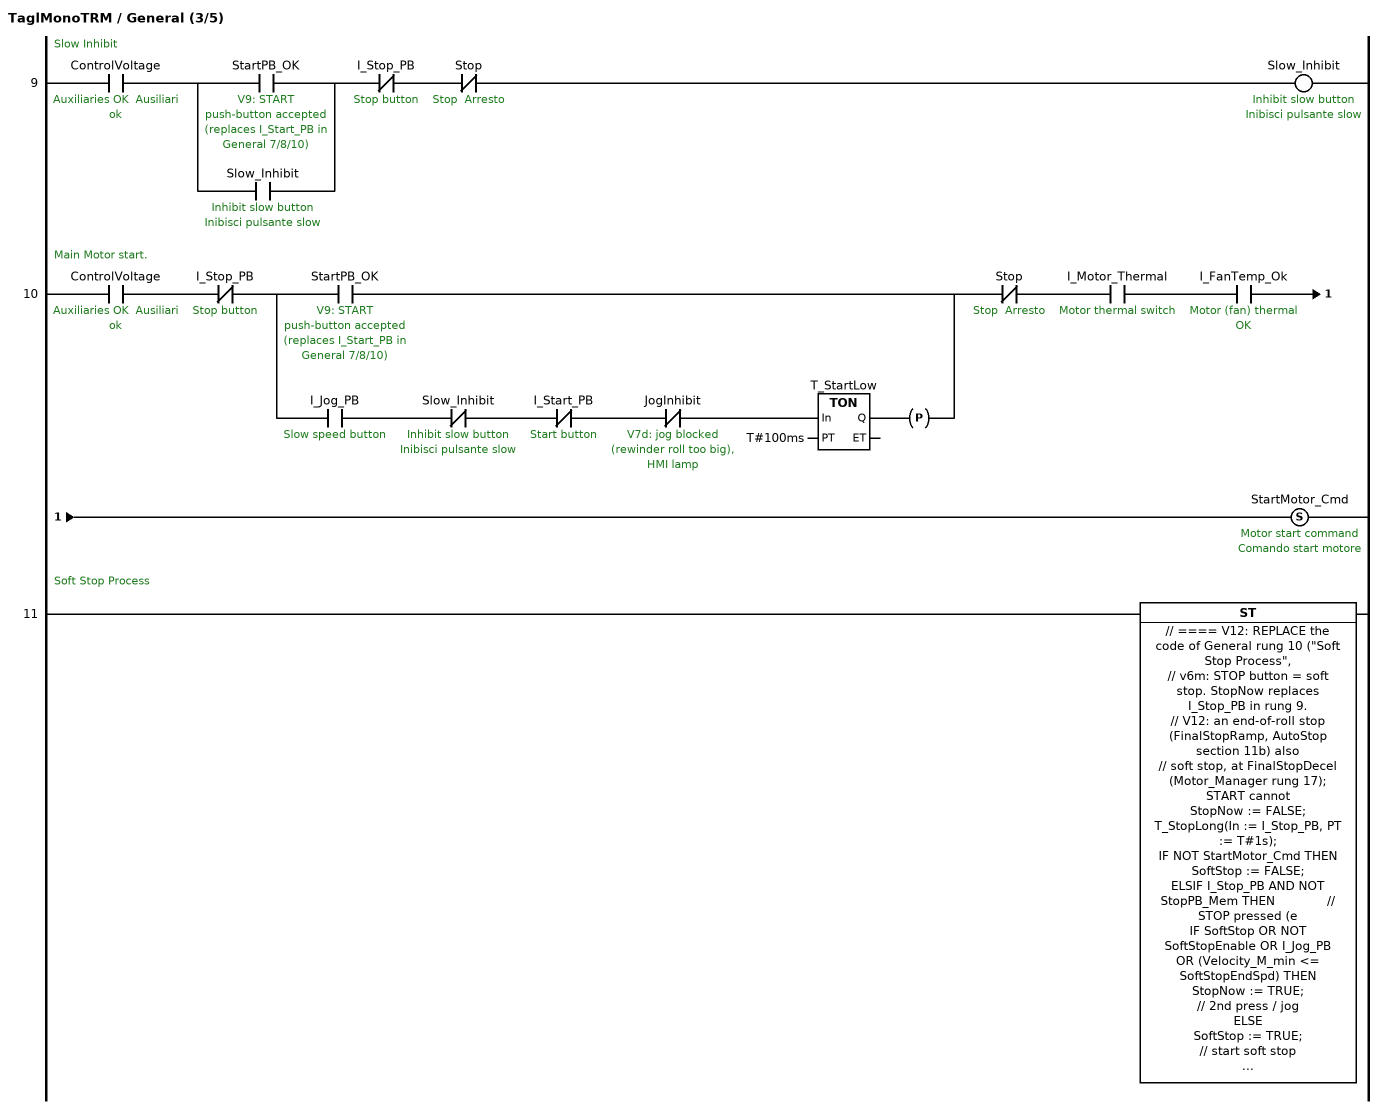
(* Rung 9: Slow Inhibit *)
Slow_Inhibit := ControlVoltage AND (StartPB_OK OR Slow_Inhibit) AND NOT I_Stop_PB AND NOT Stop;
(* Rung 10: Main Motor start. *)
T_StartLow(In := ControlVoltage AND NOT I_Stop_PB AND I_Jog_PB AND NOT Slow_Inhibit AND NOT I_Start_PB AND NOT JogInhibit, PT := T#100ms);
_e2(CLK := T_StartLow.Q);
IF ((ControlVoltage AND NOT I_Stop_PB AND StartPB_OK) OR _e2.Q) AND NOT Stop AND I_Motor_Thermal AND I_FanTemp_Ok THEN
    StartMotor_Cmd := TRUE;
END_IF;
(* Rung 11: Soft Stop Process *)
// ==== V12: REPLACE the code of General rung 10 ("Soft Stop Process", printed V9).
// v6m: STOP button = soft stop. StopNow replaces I_Stop_PB in rung 9.
// V12: an end-of-roll stop (FinalStopRamp, AutoStop section 11b) also starts the
// soft stop, at FinalStopDecel (Motor_Manager rung 17); START cannot cancel it.

StopNow := FALSE;
T_StopLong(In := I_Stop_PB, PT := T#1s);

IF NOT StartMotor_Cmd THEN
    SoftStop := FALSE;
ELSIF I_Stop_PB AND NOT StopPB_Mem THEN             // STOP pressed (edge)
	
    IF SoftStop OR NOT SoftStopEnable OR I_Jog_PB
       OR (Velocity_M_min <= SoftStopEndSpd) THEN
        StopNow := TRUE;                            // 2nd press / jog / slow / disabled
    ELSE
        SoftStop := TRUE;                           // start soft stop
    END_IF;
END_IF;

StopPB_Mem := I_Stop_PB;

IF T_StopLong.Q THEN
    StopNow := TRUE;                                // held 1 s = immediate
END_IF;

// V12: end-of-roll stop ramp (FinalStopRamp set by AutoStop section 11b)

IF FinalStopRamp AND StartMotor_Cmd AND NOT SoftStop THEN
    SoftStop := TRUE;
END_IF;

IF SoftStop AND I_Start_PB AND NOT FinalStopRamp THEN
    SoftStop := FALSE;                              // START cancels the soft stop
END_IF;

T_SoftStop(In := SoftStop, PT := T#120s);

IF SoftStop AND ((Velocity_M_min <= SoftStopEndSpd) OR T_SoftStop.Q) THEN
    StopNow := TRUE;                                // almost stopped (or timeout)
END_IF;

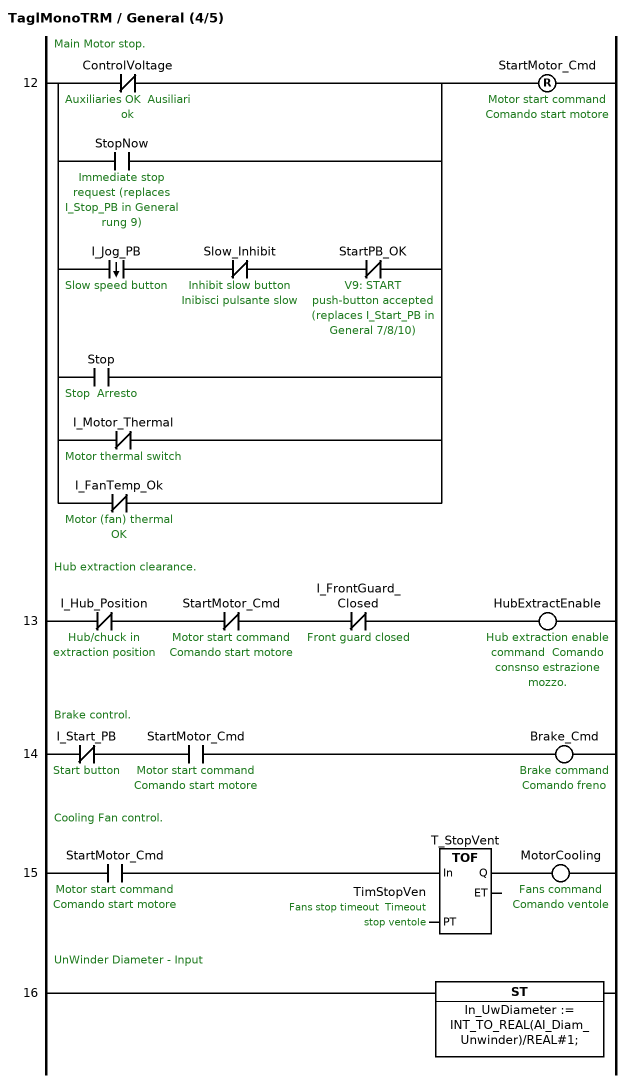
(* Rung 12: Main Motor stop. *)
_e3(CLK := I_Jog_PB);
IF NOT ControlVoltage OR StopNow OR (_e3.Q AND NOT Slow_Inhibit AND NOT StartPB_OK) OR Stop OR NOT I_Motor_Thermal OR NOT I_FanTemp_Ok THEN
    StartMotor_Cmd := FALSE;
END_IF;
(* Rung 13: Hub extraction clearance. *)
HubExtractEnable := NOT I_Hub_Position AND NOT StartMotor_Cmd AND NOT I_FrontGuard_Closed;
(* Rung 14: Brake control. *)
Brake_Cmd := NOT I_Start_PB AND StartMotor_Cmd;
(* Rung 15: Cooling Fan control. *)
T_StopVent(In := StartMotor_Cmd, PT := TimStopVen);
MotorCooling := T_StopVent.Q;
(* Rung 16: UnWinder Diameter - Input *)
In_UwDiameter := INT_TO_REAL(AI_Diam_Unwinder)/REAL#1;

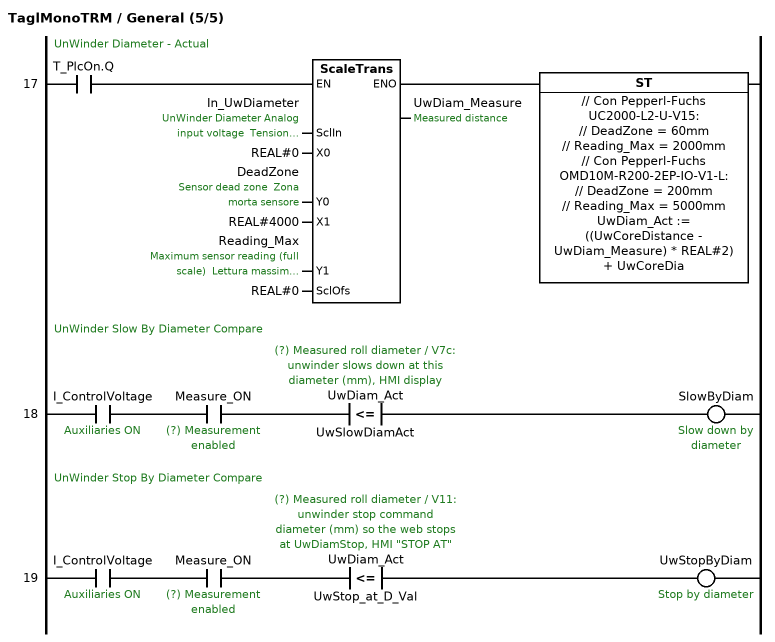
(* Rung 17: UnWinder Diameter - Actual *)
IF T_PlcOn.Q THEN
    UwDiam_Measure := ScaleTrans(SclIn := In_UwDiameter, X0 := REAL#0, Y0 := DeadZone, X1 := REAL#4000, Y1 := Reading_Max, SclOfs := REAL#0);
END_IF;
IF T_PlcOn.Q THEN
    // Con Pepperl-Fuchs UC2000-L2-U-V15:
    // DeadZone = 60mm
    // Reading_Max = 2000mm
    
    // Con Pepperl-Fuchs OMD10M-R200-2EP-IO-V1-L:
    // DeadZone = 200mm
    // Reading_Max = 5000mm
    
    UwDiam_Act := ((UwCoreDistance - UwDiam_Measure) * REAL#2) + UwCoreDiameter;
END_IF;
(* Rung 18: UnWinder Slow By Diameter Compare *)
SlowByDiam := I_ControlVoltage AND Measure_ON AND (UwDiam_Act <= UwSlowDiamAct);
(* Rung 19: UnWinder Stop By Diameter Compare *)
UwStopByDiam := I_ControlVoltage AND Measure_ON AND (UwDiam_Act <= UwStop_at_D_Val);

(* Section Motor_Manager: ladder, written here as Structured Text *)

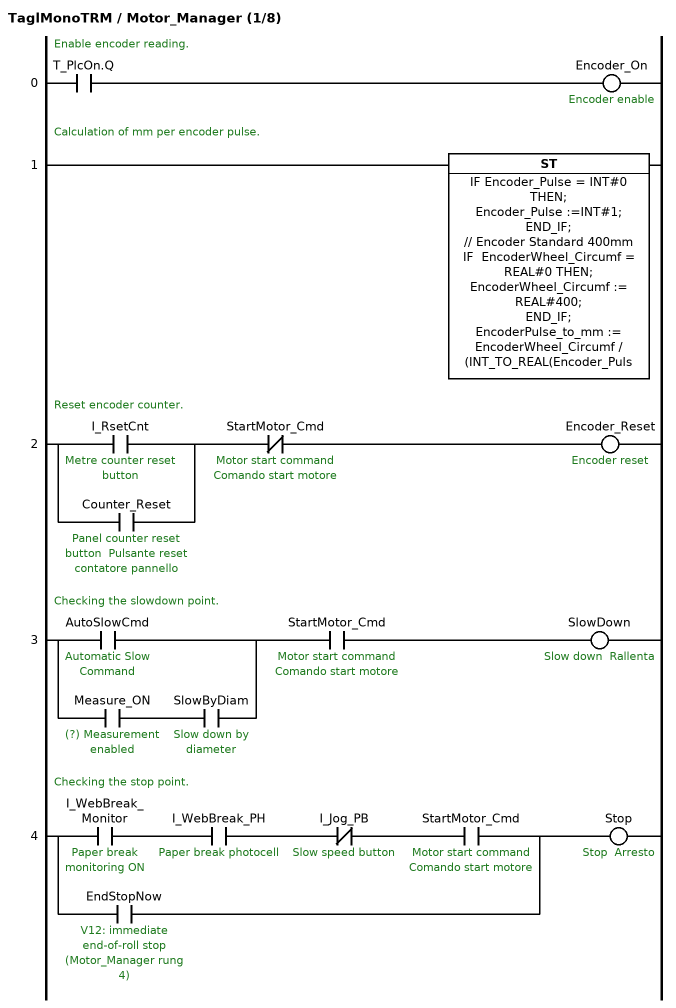
(* Rung 0: Enable encoder reading. *)
Encoder_On := T_PlcOn.Q;
(* Rung 1: Calculation of mm per encoder pulse. *)
IF Encoder_Pulse = INT#0 THEN;
	Encoder_Pulse :=INT#1;
END_IF;
// Encoder Standard 400mm
IF  EncoderWheel_Circumf = REAL#0 THEN;
	EncoderWheel_Circumf := REAL#400;
END_IF;

EncoderPulse_to_mm := EncoderWheel_Circumf / (INT_TO_REAL(Encoder_Pulse) * REAL#4);
(* Rung 2: Reset encoder counter. *)
Encoder_Reset := (I_RsetCnt OR Counter_Reset) AND NOT StartMotor_Cmd;
(* Rung 3: Checking the slowdown point. *)
SlowDown := (AutoSlowCmd OR (Measure_ON AND SlowByDiam)) AND StartMotor_Cmd;
(* Rung 4: Checking the stop point. *)
Stop := (I_WebBreak_Monitor AND I_WebBreak_PH AND NOT I_Jog_PB AND StartMotor_Cmd) OR EndStopNow;

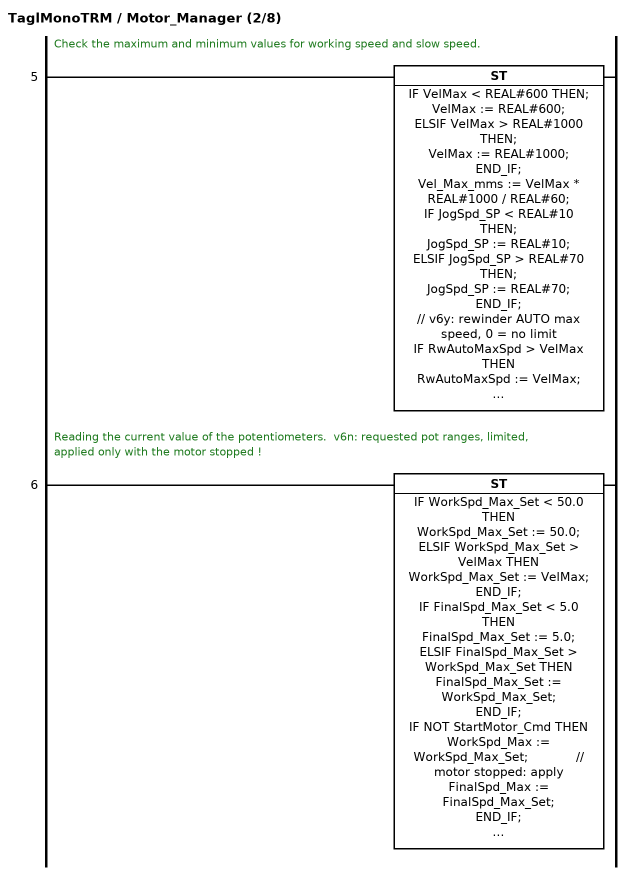
(* Rung 5: Check the maximum and minimum values ​​for working speed and slow speed. *)
IF VelMax < REAL#600 THEN;
        VelMax := REAL#600;
    ELSIF VelMax > REAL#1000 THEN;
        VelMax := REAL#1000;
END_IF;
Vel_Max_mms := VelMax * REAL#1000 / REAL#60;

IF JogSpd_SP < REAL#10 THEN;
		JogSpd_SP := REAL#10;
ELSIF JogSpd_SP > REAL#70 THEN;
	JogSpd_SP := REAL#70;
END_IF;

// v6y: rewinder AUTO max speed, 0 = no limit

IF RwAutoMaxSpd > VelMax THEN
    RwAutoMaxSpd := VelMax;
ELSIF (RwAutoMaxSpd > REAL#0) AND (RwAutoMaxSpd < REAL#50) THEN
    RwAutoMaxSpd := REAL#50;
END_IF;

IF NOT StartMotor_Cmd THEN          // taken over at standstill only
    RwAutoLimAct := RwStopEnable AND (RwAutoMaxSpd > REAL#0);
    RwAutoMaxSpdAct := RwAutoMaxSpd;
END_IF;

// ---- V7: add at the END of Motor_Manager rung 5 ("Check the maximum and minimum values...")
// ---- after the JogSpd_SP clamp, before Output_Ratio. Same style as the VelMax / JogSpd clamps.
// V7: limits on settings that stop the machine or break the auto stop if 0 / absurd

IF SpdDelta_Percent < REAL#2 THEN                  // fine band [m/min]: 0 = speed hunting
    SpdDelta_Percent := REAL#2;
ELSIF SpdDelta_Percent > REAL#15 THEN
    SpdDelta_Percent := REAL#15;
END_IF;

IF AccelTrim < REAL#0.02 THEN                      // trim ramps: 0 = no speed correction
    AccelTrim := REAL#0.02;
ELSIF AccelTrim > REAL#0.5 THEN
    AccelTrim := REAL#0.5;
END_IF;

IF DecelTrim < REAL#0.02 THEN
    DecelTrim := REAL#0.02;
ELSIF DecelTrim > REAL#0.5 THEN
    DecelTrim := REAL#0.5;
END_IF;

IF AccelCoarse < REAL#0.2 THEN                     // coarse ramps: 0 = never reaches speed
    AccelCoarse := REAL#0.2;
ELSIF AccelCoarse > REAL#4 THEN
    AccelCoarse := REAL#4;
END_IF;

IF DecelCoarse < REAL#0.2 THEN
    DecelCoarse := REAL#0.2;
ELSIF DecelCoarse > REAL#4 THEN
    DecelCoarse := REAL#4;
END_IF;

IF DecelWeb > REAL#0 THEN                          // V7 web ramps: 0 = old coarse ramp (allowed)
    IF DecelWeb < REAL#50 THEN
        DecelWeb := REAL#50;
    ELSIF DecelWeb > REAL#1000 THEN
        DecelWeb := REAL#1000;
    END_IF;
END_IF;

IF AccelWeb > REAL#0 THEN
    IF AccelWeb < REAL#50 THEN
        AccelWeb := REAL#50;
    ELSIF AccelWeb > REAL#1000 THEN
        AccelWeb := REAL#1000;
    END_IF;
END_IF;

IF SoftStopDecel > REAL#1500 THEN                  // 0 = DecelCoarse (allowed)
    SoftStopDecel := REAL#1500;
END_IF;

IF RwMaxDiam > REAL#1450 THEN                      // rewinder MECHANICAL limit [mm]
    RwMaxDiam := REAL#1450;
ELSIF RwMaxDiam < REAL#300 THEN
    RwMaxDiam := REAL#300;
END_IF;

IF RwMaxSlowFallback >= RwMaxDiam THEN             // fallback slow-down below the max
    RwMaxSlowFallback := RwMaxDiam - REAL#30;
END_IF;

// ---- V9 (V7d): add at the END of Motor_Manager rung 5, after the V7 clamps
// ---- (last lines now: RwMaxSlowFallback clamp), before Output_Ratio / Input_Ratio.
// V7d: jog / slow start button blocked on a big rewinder roll.
// RwJogMaxDiam (mm, HMI, Retain): 0 = no limit, else min 150.
// DT35 fault -> jog allowed (needed to thread / clear the machine).

IF (RwJogMaxDiam > REAL#0) AND (RwJogMaxDiam < REAL#150) THEN
    RwJogMaxDiam := REAL#150;
END_IF;

JogInhibit := (RwJogMaxDiam > REAL#0) AND (RwDiam > RwJogMaxDiam) AND NOT RwSensFault;

Output_Ratio := (VelMax * Mt_To_mm) / UINT_TO_REAL(Analog_Res); //REAL#4000;
Input_Ratio := UINT_TO_REAL(Analog_Res) / VelMax ;
(* Rung 6: Reading the current value of the potentiometers.  v6n: requested pot ranges, limited, applied only with the motor stopped ! *)
IF WorkSpd_Max_Set < 50.0 THEN
    WorkSpd_Max_Set := 50.0;
ELSIF WorkSpd_Max_Set > VelMax THEN
    WorkSpd_Max_Set := VelMax;
END_IF;

IF FinalSpd_Max_Set < 5.0 THEN
    FinalSpd_Max_Set := 5.0;
ELSIF FinalSpd_Max_Set > WorkSpd_Max_Set THEN
    FinalSpd_Max_Set := WorkSpd_Max_Set;
END_IF;

IF NOT StartMotor_Cmd THEN
    WorkSpd_Max := WorkSpd_Max_Set;            // motor stopped: apply
    FinalSpd_Max := FinalSpd_Max_Set;
END_IF;

SpdMax_Pending := (WorkSpd_Max <> WorkSpd_Max_Set)
               OR (FinalSpd_Max <> FinalSpd_Max_Set)
               OR (RwAutoLimAct <> (RwStopEnable AND (RwAutoMaxSpd > REAL#0)))
               OR (RwAutoLimAct AND (RwAutoMaxSpdAct <> RwAutoMaxSpd));

// v6i: pots scaled to their own full scale (m/min)

IF Pot1_Work_Velocity > INT#5 THEN
    Pot1_Mem := REAL_TO_INT(INT_TO_REAL(Pot1_Work_Velocity) * WorkSpd_Max / VelMax);
ELSE
    Pot1_Mem := INT#0;
END_IF;

IF Pot2_Slow_Velocity > INT#5 THEN
    Pot2_Mem := REAL_TO_INT(INT_TO_REAL(Pot2_Slow_Velocity) * FinalSpd_Max / VelMax);
ELSE
    Pot2_Mem := INT#0;
END_IF;

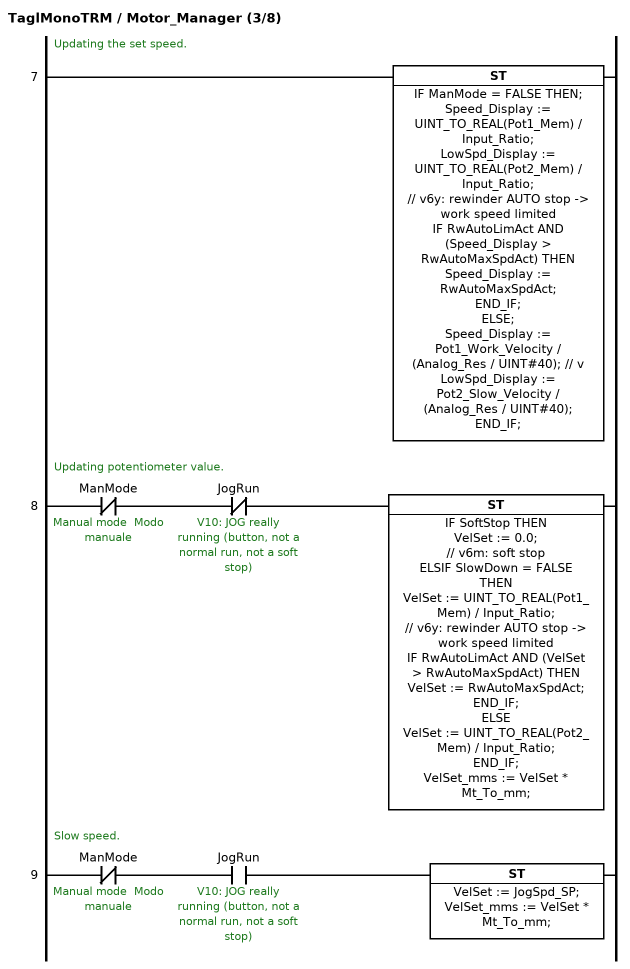
(* Rung 7: Updating the set speed. *)
IF ManMode = FALSE THEN;
		
		Speed_Display := UINT_TO_REAL(Pot1_Mem) / Input_Ratio;
		LowSpd_Display := UINT_TO_REAL(Pot2_Mem) / Input_Ratio;
			
     // v6y: rewinder AUTO stop -> work speed limited
	
     IF RwAutoLimAct AND (Speed_Display > RwAutoMaxSpdAct) THEN
         Speed_Display := RwAutoMaxSpdAct;
     END_IF;
				
ELSE;
    Speed_Display := Pot1_Work_Velocity / (Analog_Res / UINT#40); // v6i: raw pot, %
    LowSpd_Display := Pot2_Slow_Velocity / (Analog_Res / UINT#40);
	
END_IF;
(* Rung 8: Updating potentiometer value. *)
IF NOT ManMode AND NOT JogRun THEN
    IF SoftStop THEN
        VelSet := 0.0;                                  // v6m: soft stop
    ELSIF SlowDown = FALSE  THEN
        VelSet := UINT_TO_REAL(Pot1_Mem) / Input_Ratio;
    	
        // v6y: rewinder AUTO stop -> work speed limited
    	
        IF RwAutoLimAct AND (VelSet > RwAutoMaxSpdAct) THEN
            VelSet := RwAutoMaxSpdAct;
        END_IF;
    	
    ELSE
        VelSet := UINT_TO_REAL(Pot2_Mem) / Input_Ratio;
    END_IF;
    
    VelSet_mms := VelSet * Mt_To_mm;
END_IF;
(* Rung 9: Slow speed. *)
IF NOT ManMode AND JogRun THEN
    VelSet := JogSpd_SP;
    VelSet_mms := VelSet * Mt_To_mm;
END_IF;

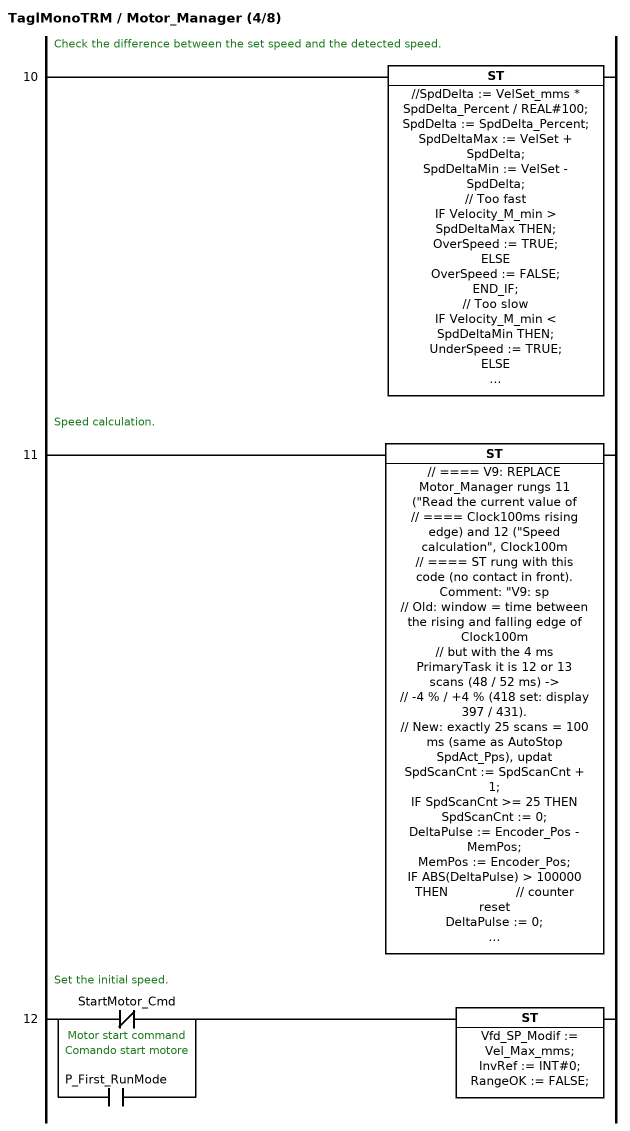
(* Rung 10: Check the difference between the set speed and the detected speed. *)
//SpdDelta := VelSet_mms * SpdDelta_Percent / REAL#100;

SpdDelta := SpdDelta_Percent;
SpdDeltaMax := VelSet + SpdDelta;
SpdDeltaMin := VelSet - SpdDelta;

// Too fast

IF Velocity_M_min > SpdDeltaMax THEN;
		OverSpeed := TRUE;
	ELSE
		OverSpeed := FALSE;
END_IF;

// Too slow

IF Velocity_M_min < SpdDeltaMin THEN;
		UnderSpeed := TRUE;
	ELSE
		UnderSpeed := FALSE;
END_IF;
(* Rung 11: Speed ​​calculation. *)
// ==== V9: REPLACE Motor_Manager rungs 11 ("Read the current value of the encoder", MOVE on
// ==== Clock100ms rising edge) and 12 ("Speed calculation", Clock100ms falling edge) by ONE
// ==== ST rung with this code (no contact in front). Comment: "V9: speed over exactly 100 ms".
// Old: window = time between the rising and falling edge of Clock100ms, assumed 50 ms,
// but with the 4 ms PrimaryTask it is 12 or 13 scans (48 / 52 ms) -> the speed jumps
// -4 % / +4 % (418 set: display 397 / 431).
// New: exactly 25 scans = 100 ms (same as AutoStop SpdAct_Pps), updated 10 times/s.

SpdScanCnt := SpdScanCnt + 1;

IF SpdScanCnt >= 25 THEN
    SpdScanCnt := 0;
    DeltaPulse := Encoder_Pos - MemPos;
    MemPos := Encoder_Pos;
	
    IF ABS(DeltaPulse) > 100000 THEN                 // counter reset (Encoder_Reset)
        DeltaPulse := 0;
    END_IF;
	
    Velocity := DINT_TO_REAL(DeltaPulse) * EncoderPulse_to_mm * REAL#10;   // mm/s
    Velocity_M_min := Velocity / Mt_To_mm;
END_IF;
(* Rung 12: Set the initial speed. *)
IF NOT StartMotor_Cmd OR P_First_RunMode THEN
    Vfd_SP_Modif := Vel_Max_mms;
    InvRef := INT#0;
    RangeOK := FALSE;
END_IF;

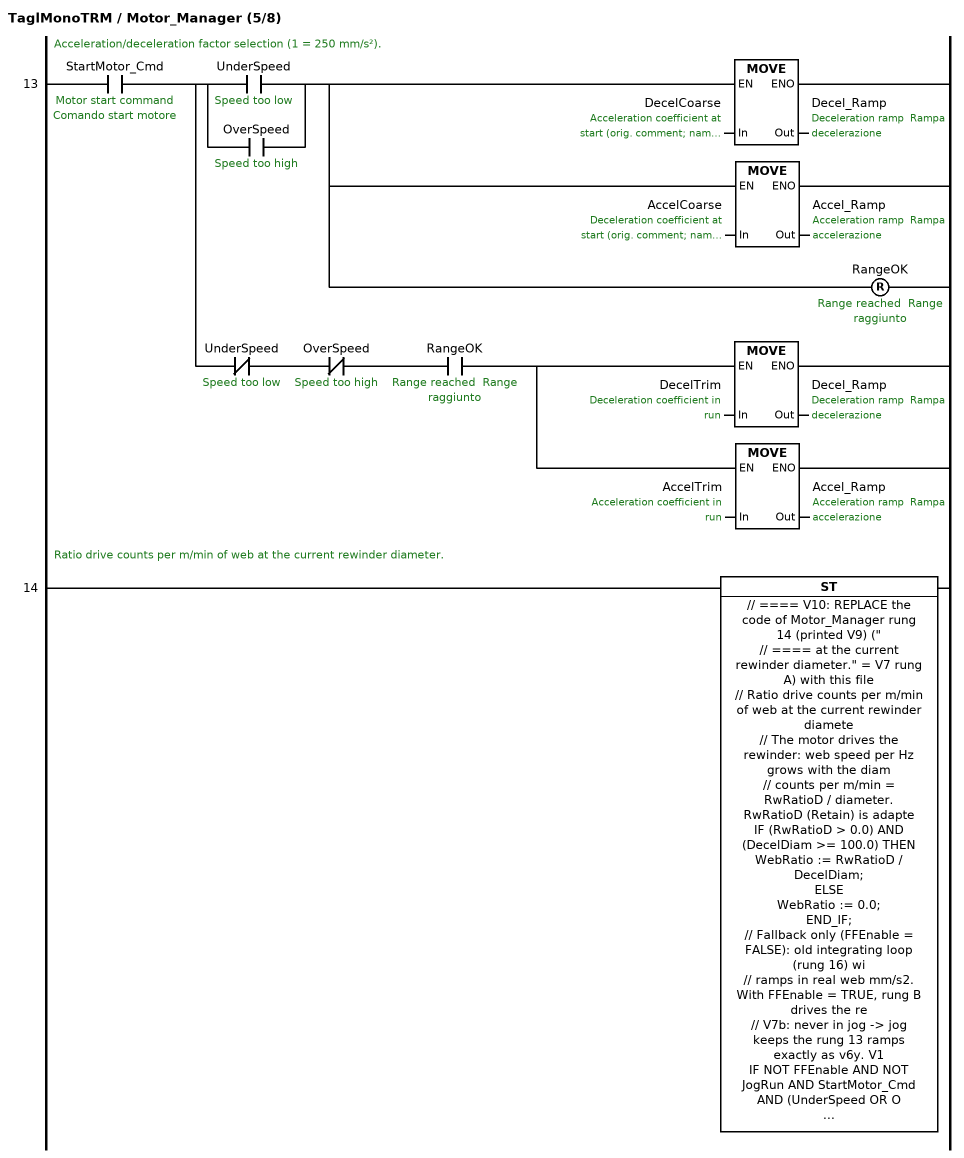
(* Rung 13: Acceleration/deceleration factor selection (1 = 250 mm/s²). *)
IF StartMotor_Cmd AND (UnderSpeed OR OverSpeed) THEN
    Decel_Ramp := DecelCoarse;
    Accel_Ramp := AccelCoarse;
    RangeOK := FALSE;
END_IF;
_p4 := StartMotor_Cmd AND NOT UnderSpeed AND NOT OverSpeed AND RangeOK;
IF _p4 THEN
    Decel_Ramp := DecelTrim;
    Accel_Ramp := AccelTrim;
END_IF;
(* Rung 14: Ratio drive counts per m/min of web at the current rewinder diameter. *)
// ==== V10: REPLACE the code of Motor_Manager rung 14 (printed V9) ("Ratio drive counts per m/min of web
// ==== at the current rewinder diameter." = V7 rung A) with this file. (V7b jog line inside.)
// Ratio drive counts per m/min of web at the current rewinder diameter.
// The motor drives the rewinder: web speed per Hz grows with the diameter, so
// counts per m/min = RwRatioD / diameter. RwRatioD (Retain) is adapted by rung B.

IF (RwRatioD > 0.0) AND (DecelDiam >= 100.0) THEN
    WebRatio := RwRatioD / DecelDiam;
ELSE
    WebRatio := 0.0;
END_IF;

// Fallback only (FFEnable = FALSE): old integrating loop (rung 16) with the coarse
// ramps in real web mm/s2. With FFEnable = TRUE, rung B drives the reference.
// V7b: never in jog -> jog keeps the rung 13 ramps exactly as v6y. V10: JogRun (jog really running).

IF NOT FFEnable AND NOT JogRun AND StartMotor_Cmd AND (UnderSpeed OR OverSpeed)
   AND (WebRatio > 0.0) THEN
   
    IF DecelWeb > 0.0 THEN
        Decel_Ramp := DecelWeb * 0.06 * WebRatio * Vel_Max_mms / 1000000.0;
        IF Decel_Ramp > 8.0 THEN
            Decel_Ramp := 8.0;
        END_IF;
    END_IF;
	
    IF AccelWeb > 0.0 THEN
        Accel_Ramp := AccelWeb * 0.06 * WebRatio * Vel_Max_mms / 1000000.0;
		
        IF Accel_Ramp > 8.0 THEN
            Accel_Ramp := 8.0;
        END_IF;
    END_IF;
END_IF;

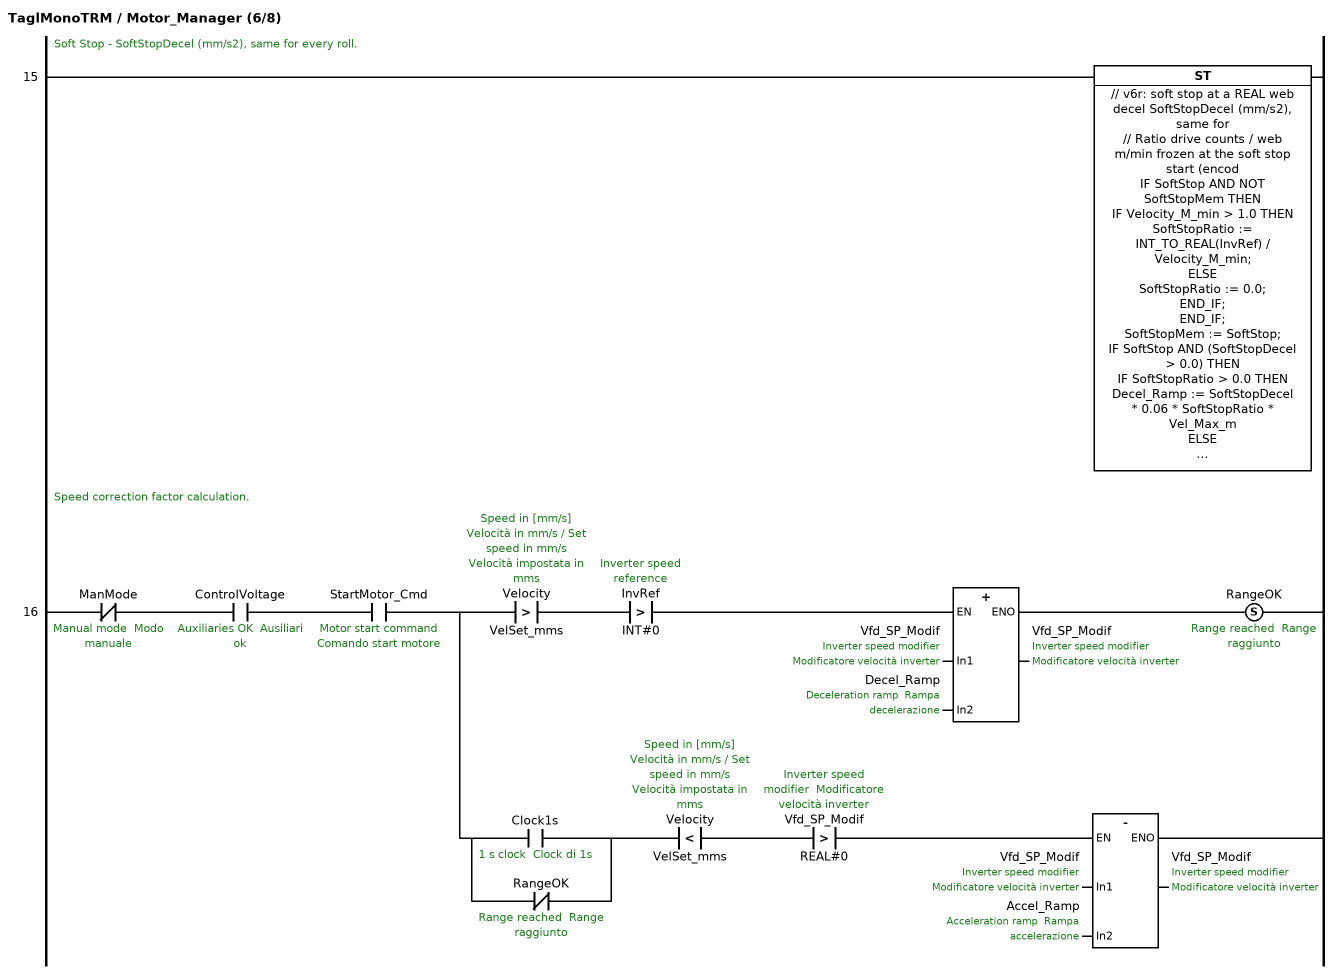
(* Rung 15: Soft Stop - SoftStopDecel (mm/s2), same for every roll. *)
// v6r: soft stop at a REAL web decel SoftStopDecel (mm/s2), same for every roll.
// Ratio drive counts / web m/min frozen at the soft stop start (encoder = exact).

IF SoftStop AND NOT SoftStopMem THEN
    IF Velocity_M_min > 1.0 THEN
        SoftStopRatio := INT_TO_REAL(InvRef) / Velocity_M_min;
    ELSE
        SoftStopRatio := 0.0;
    END_IF;
END_IF;

SoftStopMem := SoftStop;

IF SoftStop AND (SoftStopDecel > 0.0) THEN
    IF SoftStopRatio > 0.0 THEN
        Decel_Ramp := SoftStopDecel * 0.06 * SoftStopRatio * Vel_Max_mms / 1000000.0;
    ELSE
        Decel_Ramp := SoftStopDecel / 250.0;            // fallback (old v6m behaviour)
    END_IF;
	
    IF Decel_Ramp > 8.0 THEN
        Decel_Ramp := 8.0;                              // max 9 Hz/s asked from the PLC
    END_IF;
END_IF;
(* Rung 16: Speed ​​correction factor calculation. *)
_p5 := NOT ManMode AND ControlVoltage AND StartMotor_Cmd;
IF _p5 AND (Velocity > VelSet_mms) AND (InvRef > INT#0) THEN
    Vfd_SP_Modif := Vfd_SP_Modif + Decel_Ramp;
    RangeOK := TRUE;
END_IF;
IF _p5 AND (Clock1s OR NOT RangeOK) AND (Velocity < VelSet_mms) AND (Vfd_SP_Modif > REAL#0) THEN
    Vfd_SP_Modif := Vfd_SP_Modif - Accel_Ramp;
END_IF;

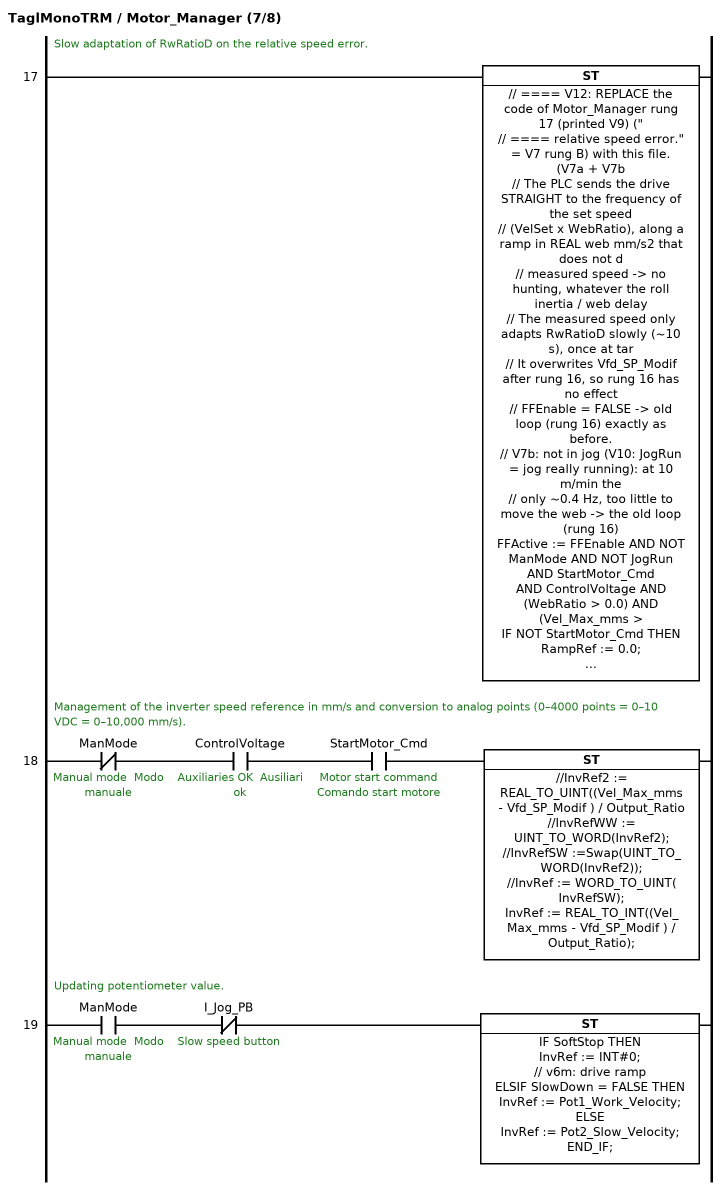
(* Rung 17: Slow adaptation of RwRatioD on the relative speed error. *)
// ==== V12: REPLACE the code of Motor_Manager rung 17 (printed V9) ("Slow adaptation of RwRatioD on the
// ==== relative speed error." = V7 rung B) with this file. (V7a + V7b + V7f + V9 + V10 + V12 inside.)
// The PLC sends the drive STRAIGHT to the frequency of the set speed
// (VelSet x WebRatio), along a ramp in REAL web mm/s2 that does not depend on the
// measured speed -> no hunting, whatever the roll inertia / web delay.
// The measured speed only adapts RwRatioD slowly (~10 s), once at target.
// It overwrites Vfd_SP_Modif after rung 16, so rung 16 has no effect in AUTO.
// FFEnable = FALSE -> old loop (rung 16) exactly as before.
// V7b: not in jog (V10: JogRun = jog really running): at 10 m/min the feed-forward gives
// only ~0.4 Hz, too little to move the web -> the old loop (rung 16) runs the jog.

FFActive := FFEnable AND NOT ManMode AND NOT JogRun AND StartMotor_Cmd
            AND ControlVoltage AND (WebRatio > 0.0) AND (Vel_Max_mms > 0.0);

IF NOT StartMotor_Cmd THEN
    RampRef := 0.0;
    FFRate := 0.0;
    FFSteadyTicks := 0;
    FFSlowAcc := FALSE;
END_IF;

// V9: START during a soft stop: the decel flattens and the speed is HELD
// (SpdHold, HMI lamp) until START is pushed AGAIN -> gentle ramp up at
// SoftCancelAccel (mm/s2) to the set speed. The hold only blocks speeding up:
// a lower target (pot down, auto slow-down, RwAutoMaxSpd) still slows down.
// STOP during the hold = new soft stop (General rung 9).

IF (SoftCancelAccel > 0.0) AND (SoftCancelAccel < 20.0) THEN
    SoftCancelAccel := 20.0;
ELSIF SoftCancelAccel > 1000.0 THEN
    SoftCancelAccel := 1000.0;
END_IF;

FFStartEdge := I_Start_PB AND NOT FFStartMem;
FFStartMem := I_Start_PB;

IF FFSoftMem AND NOT SoftStop AND StartMotor_Cmd AND FFActive THEN   // soft stop cancelled
    SpdHold := TRUE;
    FFSlowAcc := FALSE;
ELSIF SpdHold AND FFStartEdge THEN                       // 2nd START: resume
    SpdHold := FALSE;
    FFSlowAcc := TRUE;
END_IF;

IF SoftStop OR NOT StartMotor_Cmd OR NOT FFActive THEN    // FFEnable OFF: old loop
    SpdHold := FALSE;
    FFSlowAcc := FALSE;
END_IF;

FFSoftMem := SoftStop;

// V7f: S-curve time (s), 0 = off, max 2 s

IF SCurveTime < 0.0 THEN
    SCurveTime := 0.0;
ELSIF SCurveTime > 2.0 THEN
    SCurveTime := 2.0;
END_IF;

IF FFActive THEN
    IF NOT FFWasActive THEN
        RampRef := Vel_Max_mms - Vfd_SP_Modif;          // bumpless start / switch-over
        FFRate := 0.0;
    END_IF;

    // Target reference (mm/s of the 0..10 V scale) for the set speed	
    FFTarget := VelSet * WebRatio * Output_Ratio;
	
    IF FFTarget > Vel_Max_mms THEN
        FFTarget := Vel_Max_mms;
    ELSIF FFTarget < 0.0 THEN
        FFTarget := 0.0;
    END_IF;

    // Tension: hold at TensWaitSpd until the T-one reports tension (I_T_one_TensionOK)
	
    IF TensWait AND (VelSet > TensWaitSpd) THEN
        FFTarget := TensWaitSpd * WebRatio * Output_Ratio;
    END_IF;

    // V9: hold after a cancelled soft stop (the S-curve flattens it smoothly):
    // never above the present reference, lower targets still allowed
	
    IF SpdHold THEN
        IF FFTarget > RampRef THEN
            FFTarget := RampRef;
        END_IF;
		
    ELSIF FFSlowAcc AND (ABS(FFTarget - RampRef) <= FFTarget * 0.005 + 2.0) THEN
        FFSlowAcc := FALSE;                              // back at the set speed
    END_IF;

    // Ramp steps per 4 ms scan: web mm/s2 -> reference mm/s per scan
	
    IF FFSlowAcc AND (SoftCancelAccel > 0.0) THEN
        StepAcc := SoftCancelAccel * 0.06 * WebRatio * Vel_Max_mms / 1000000.0;   // V9
    ELSIF AccelWeb > 0.0 THEN
        StepAcc := AccelWeb * 0.06 * WebRatio * Vel_Max_mms / 1000000.0;
    ELSE
        StepAcc := AccelCoarse;
    END_IF;
	
    IF SoftStop AND FinalStopRamp AND (FinalStopDecel > 0.0) THEN
        StepDec := FinalStopDecel * 0.06 * WebRatio * Vel_Max_mms / 1000000.0;   // V12 end-of-roll
    ELSIF SoftStop AND (SoftStopDecel > 0.0) THEN
        StepDec := SoftStopDecel * 0.06 * WebRatio * Vel_Max_mms / 1000000.0;
    ELSIF DecelWeb > 0.0 THEN
        StepDec := DecelWeb * 0.06 * WebRatio * Vel_Max_mms / 1000000.0;
    ELSE
        StepDec := DecelCoarse;
    END_IF;
	
    IF StepAcc > 8.0 THEN
        StepAcc := 8.0;
    END_IF;
	
    IF StepDec > 8.0 THEN
        StepDec := 8.0;
    END_IF;

    // Ramp generator
    // V7f: S-curve. FFRate (reference per scan) changes at most FFJerk per scan,
    // so the full ramp is reached after SCurveTime (s) and is rounded off the
    // same way before the target -> the T-one / brake air can follow.
    // SCurveTime = 0 -> plain linear ramp as V7a.
	
    IF SCurveTime > 0.0 THEN
        IF (FFRate > 0.0) OR ((FFRate = 0.0) AND (FFTarget > RampRef)) THEN
            FFJerk := StepAcc * 0.004 / SCurveTime;
        ELSE
            FFJerk := StepDec * 0.004 / SCurveTime;
        END_IF;
		
        // rate allowed so that it can still fall to 0 at the target
        // (no MIN(), argument in a REAL variable first: Sysmac data type rules,
        //  same pattern as SqrtArg / SQRT(SqrtArg) in AutoStop)
		
        IF FFTarget >= RampRef THEN
            FFSqrtArg := REAL#2.0 * FFJerk * (FFTarget - RampRef);
            FFRateSet := SQRT(FFSqrtArg);
			
            IF FFRateSet > StepAcc THEN
                FFRateSet := StepAcc;
            END_IF;
        ELSE
            FFSqrtArg := REAL#2.0 * FFJerk * (RampRef - FFTarget);
            FFRateSet := SQRT(FFSqrtArg);
			
            IF FFRateSet > StepDec THEN
                FFRateSet := StepDec;
            END_IF;
			
            FFRateSet := -FFRateSet;
        END_IF;
		
        IF FFRateSet > FFRate + FFJerk THEN
            FFRate := FFRate + FFJerk;
        ELSIF FFRateSet < FFRate - FFJerk THEN
            FFRate := FFRate - FFJerk;
        ELSE
            FFRate := FFRateSet;
        END_IF;
		
        RampRef := RampRef + FFRate;
		
        IF (ABS(FFTarget - RampRef) <= 3.0) AND (ABS(FFRate) <= 2.0 * FFJerk) THEN
            RampRef := FFTarget;                         // at target (pot noise)
            FFRate := 0.0;
        END_IF;
    ELSE
        FFRate := 0.0;
		
        IF RampRef < FFTarget - StepAcc THEN
            RampRef := RampRef + StepAcc;
        ELSIF RampRef > FFTarget + StepDec THEN
            RampRef := RampRef - StepDec;
        ELSE
            RampRef := FFTarget;                         // at target
        END_IF;
    END_IF;
	
    // V7a: "at target" = within 0.5 % of the target (the pot and RwDiam noise
    // move FFTarget by a few counts every scan -> the counter never reached 500)
	
    IF (ABS(FFTarget - RampRef) <= FFTarget * 0.005 + 2.0)
       AND NOT SpdHold AND NOT FFSlowAcc THEN            // V9: not during the hold
	   
        IF FFSteadyTicks < 30000 THEN
            FFSteadyTicks := FFSteadyTicks + 1;
        END_IF;
    ELSE
        FFSteadyTicks := 0;
    END_IF;

    // Slow adaptation of RwRatioD on the relative speed error (2 s after the
    // target is reached, not at the 60 Hz limit, not during soft stop / jog)
	
    IF (FFSteadyTicks >= 500) AND NOT SoftStop AND NOT JogRun
       AND (VelSet > 15.0) AND (Velocity_M_min > 10.0) AND NOT RwSensFault
       AND (FFTarget < Vel_Max_mms * 0.98) THEN
        FFErr := (VelSet - Velocity_M_min) / VelSet;
		
        IF FFErr > 0.05 THEN
            FFErr := 0.05;
        ELSIF FFErr < -0.05 THEN
            FFErr := -0.05;
        END_IF;
		
        IF ABS(FFErr) > 0.003 THEN                       // dead band 0.3 % (encoder noise)
            RwRatioD := RwRatioD * (1.0 + 0.0004 * FFErr);  // ~10 s time constant
        END_IF;
		
        IF RwRatioD < 1000.0 THEN
            RwRatioD := 1000.0;
        ELSIF RwRatioD > 8000.0 THEN
            RwRatioD := 8000.0;
        END_IF;
    END_IF;

    Vfd_SP_Modif := Vel_Max_mms - RampRef;               // rung 17 -> InvRef
END_IF;

FFWasActive := FFActive;

// V7f: T-one decel signal (for a T-one "stop / boost" input, spare PLC output):
// ON while the feed-forward ramps down (more than 1 % above the target, so the
// slow drift of the target with the diameter does not pulse it) or soft stop.

TOneDecel := (FFActive AND (RampRef - FFTarget > FFTarget * 0.01 + 5.0))
             OR (SoftStop AND StartMotor_Cmd);
(* Rung 18: Management of the inverter speed reference in mm/s and conversion to analog points (0–4000 points = 0–10 VDC = 0–10,000 mm/s). *)
IF NOT ManMode AND ControlVoltage AND StartMotor_Cmd THEN
    //InvRef2 := REAL_TO_UINT((Vel_Max_mms - Vfd_SP_Modif ) / Output_Ratio);
    //InvRefWW := UINT_TO_WORD(InvRef2);
    //InvRefSW :=Swap(UINT_TO_WORD(InvRef2));
    //InvRef := WORD_TO_UINT(InvRefSW);
    
    InvRef := REAL_TO_INT((Vel_Max_mms - Vfd_SP_Modif ) / Output_Ratio);
END_IF;
(* Rung 19: Updating potentiometer value. *)
IF ManMode AND NOT I_Jog_PB THEN
    IF SoftStop THEN
        InvRef := INT#0;                                // v6m: drive ramps down on its own
    ELSIF SlowDown = FALSE THEN
        InvRef := Pot1_Work_Velocity;
    ELSE
        InvRef := Pot2_Slow_Velocity;
    END_IF;
END_IF;

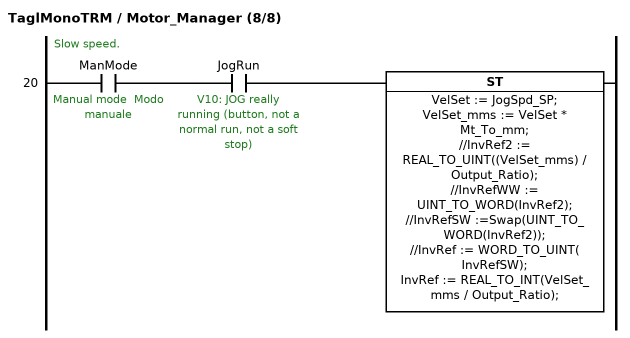
(* Rung 20: Slow speed. *)
IF ManMode AND JogRun THEN
    VelSet := JogSpd_SP;
    VelSet_mms := VelSet * Mt_To_mm;
    
    //InvRef2 := REAL_TO_UINT((VelSet_mms) / Output_Ratio);
    //InvRefWW := UINT_TO_WORD(InvRef2);
    //InvRefSW :=Swap(UINT_TO_WORD(InvRef2));
    //InvRef := WORD_TO_UINT(InvRefSW);
    
    InvRef := REAL_TO_INT(VelSet_mms / Output_Ratio);
END_IF;

(* Section OverRider_Manager: ladder, written here as Structured Text *)

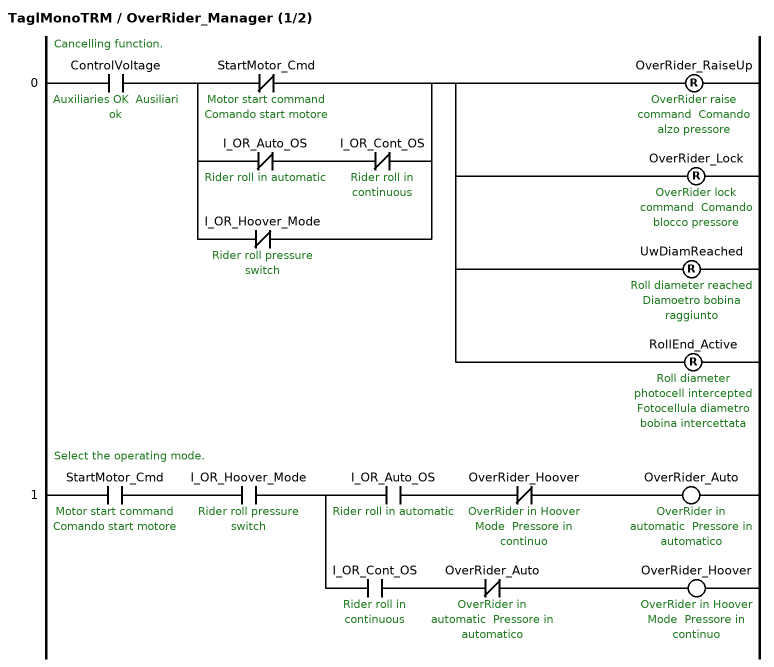
(* Rung 0: Cancelling function. *)
_p6 := ControlVoltage AND (NOT StartMotor_Cmd OR (NOT I_OR_Auto_OS AND NOT I_OR_Cont_OS) OR NOT I_OR_Hoover_Mode);
IF _p6 THEN
    OverRider_RaiseUp := FALSE;
    OverRider_Lock := FALSE;
    UwDiamReached := FALSE;
    RollEnd_Active := FALSE;
END_IF;
(* Rung 1: Select the operating mode. *)
OverRider_Auto := StartMotor_Cmd AND I_OR_Hoover_Mode AND I_OR_Auto_OS AND NOT OverRider_Hoover;
OverRider_Hoover := StartMotor_Cmd AND I_OR_Hoover_Mode AND I_OR_Cont_OS AND NOT OverRider_Auto;

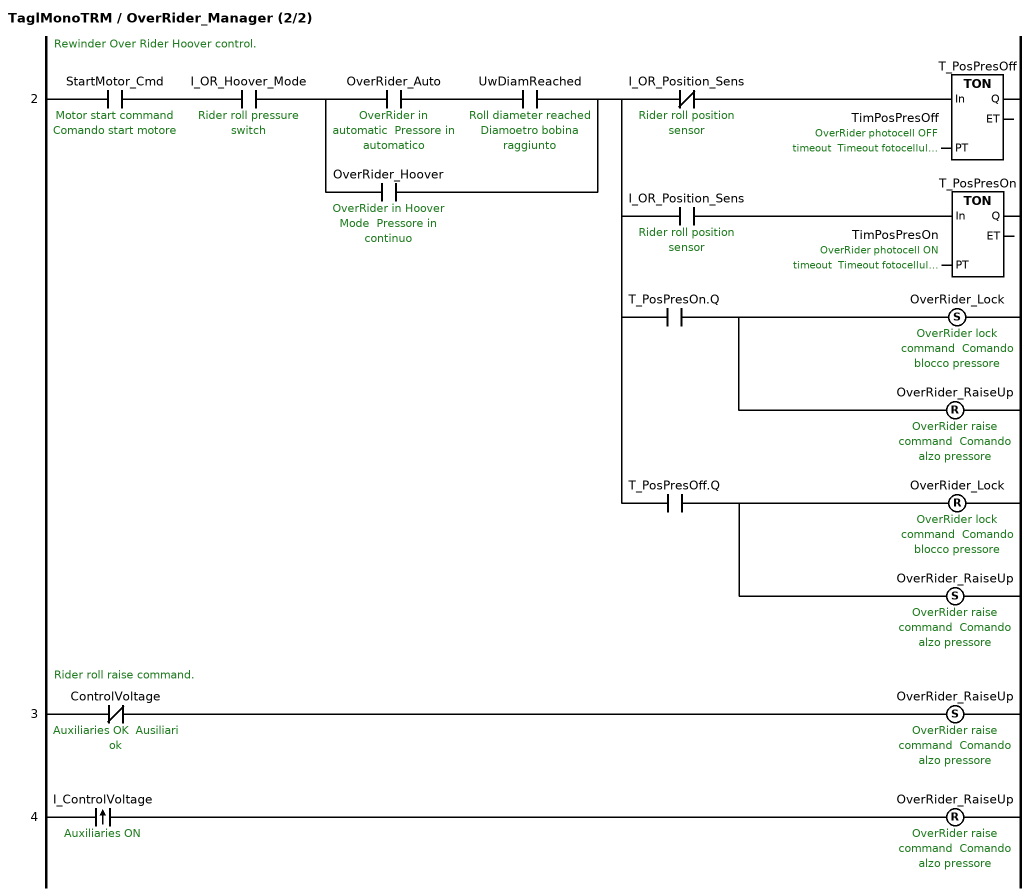
(* Rung 2: Rewinder Over Rider Hoover control. *)
_p7 := StartMotor_Cmd AND I_OR_Hoover_Mode AND ((OverRider_Auto AND UwDiamReached) OR OverRider_Hoover);
T_PosPresOff(In := _p7 AND NOT I_OR_Position_Sens, PT := TimPosPresOff);
T_PosPresOn(In := _p7 AND I_OR_Position_Sens, PT := TimPosPresOn);
IF _p7 AND T_PosPresOn.Q THEN
    OverRider_Lock := TRUE;
    OverRider_RaiseUp := FALSE;
END_IF;
IF _p7 AND T_PosPresOff.Q THEN
    OverRider_Lock := FALSE;
    OverRider_RaiseUp := TRUE;
END_IF;
(* Rung 3: Rider roll raise command. *)
IF NOT ControlVoltage THEN OverRider_RaiseUp := TRUE; END_IF;
(* Rung 4 *)
_e8(CLK := I_ControlVoltage);
IF _e8.Q THEN OverRider_RaiseUp := FALSE; END_IF;

(* Section Console: ladder, written here as Structured Text *)

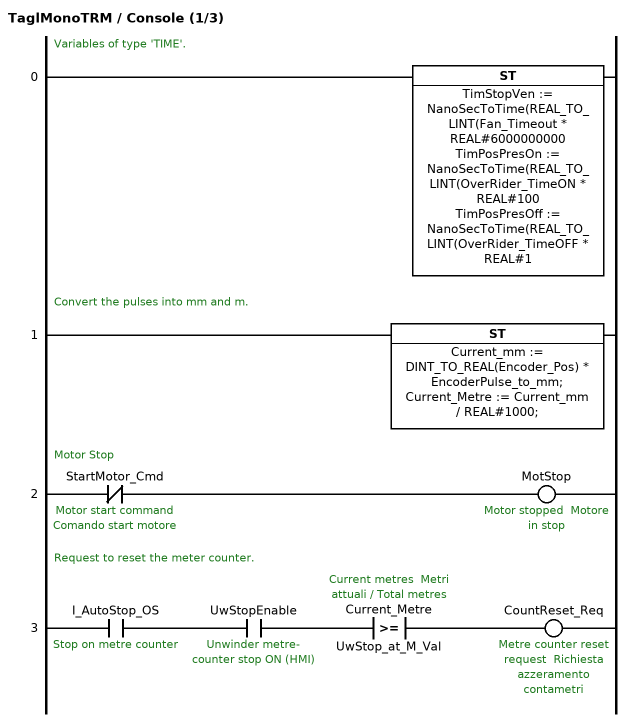
(* Rung 0: Variables of type 'TIME'. *)
TimStopVen := NanoSecToTime(REAL_TO_LINT(Fan_Timeout * REAL#60000000000));
TimPosPresOn := NanoSecToTime(REAL_TO_LINT(OverRider_TimeON * REAL#1000000000));
TimPosPresOff := NanoSecToTime(REAL_TO_LINT(OverRider_TimeOFF * REAL#1000000000));
(* Rung 1: Convert the pulses into mm and m. *)
Current_mm := DINT_TO_REAL(Encoder_Pos) * EncoderPulse_to_mm;
Current_Metre := Current_mm / REAL#1000;
(* Rung 2: Motor Stop *)
MotStop := NOT StartMotor_Cmd;
(* Rung 3: Request to reset the meter counter. *)
CountReset_Req := I_AutoStop_OS AND UwStopEnable AND (Current_Metre >= UwStop_at_M_Val);

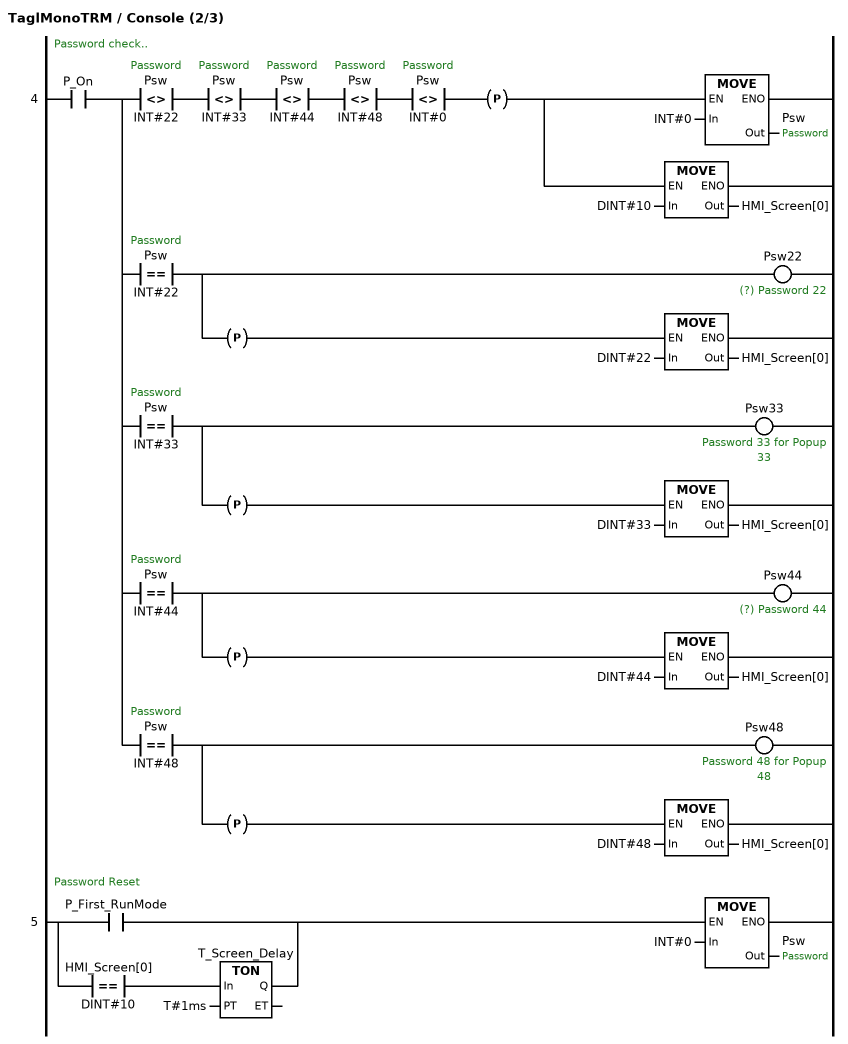
(* Rung 4: Password check.. *)
_e9(CLK := P_On AND (Psw <> INT#22) AND (Psw <> INT#33) AND (Psw <> INT#44) AND (Psw <> INT#48) AND (Psw <> INT#0));
IF _e9.Q THEN
    Psw := INT#0;
    HMI_Screen[0] := DINT#10;
END_IF;
Psw22 := P_On AND (Psw = INT#22);
_e10(CLK := P_On AND (Psw = INT#22));
IF _e10.Q THEN HMI_Screen[0] := DINT#22; END_IF;
Psw33 := P_On AND (Psw = INT#33);
_e11(CLK := P_On AND (Psw = INT#33));
IF _e11.Q THEN HMI_Screen[0] := DINT#33; END_IF;
Psw44 := P_On AND (Psw = INT#44);
_e12(CLK := P_On AND (Psw = INT#44));
IF _e12.Q THEN HMI_Screen[0] := DINT#44; END_IF;
Psw48 := P_On AND (Psw = INT#48);
_e13(CLK := P_On AND (Psw = INT#48));
IF _e13.Q THEN HMI_Screen[0] := DINT#48; END_IF;
(* Rung 5: Password Reset *)
T_Screen_Delay(In := HMI_Screen[0] = DINT#10, PT := T#1ms);
IF P_First_RunMode OR T_Screen_Delay.Q THEN Psw := INT#0; END_IF;

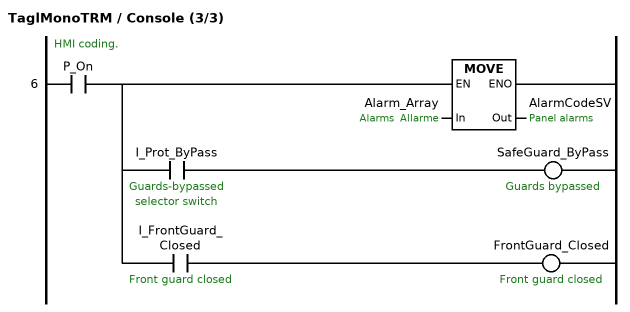
(* Rung 6: HMI coding. *)
IF P_On THEN AlarmCodeSV := Alarm_Array; END_IF;
SafeGuard_ByPass := P_On AND I_Prot_ByPass;
FrontGuard_Closed := P_On AND I_FrontGuard_Closed;

(* Section Alarms: ladder, written here as Structured Text *)

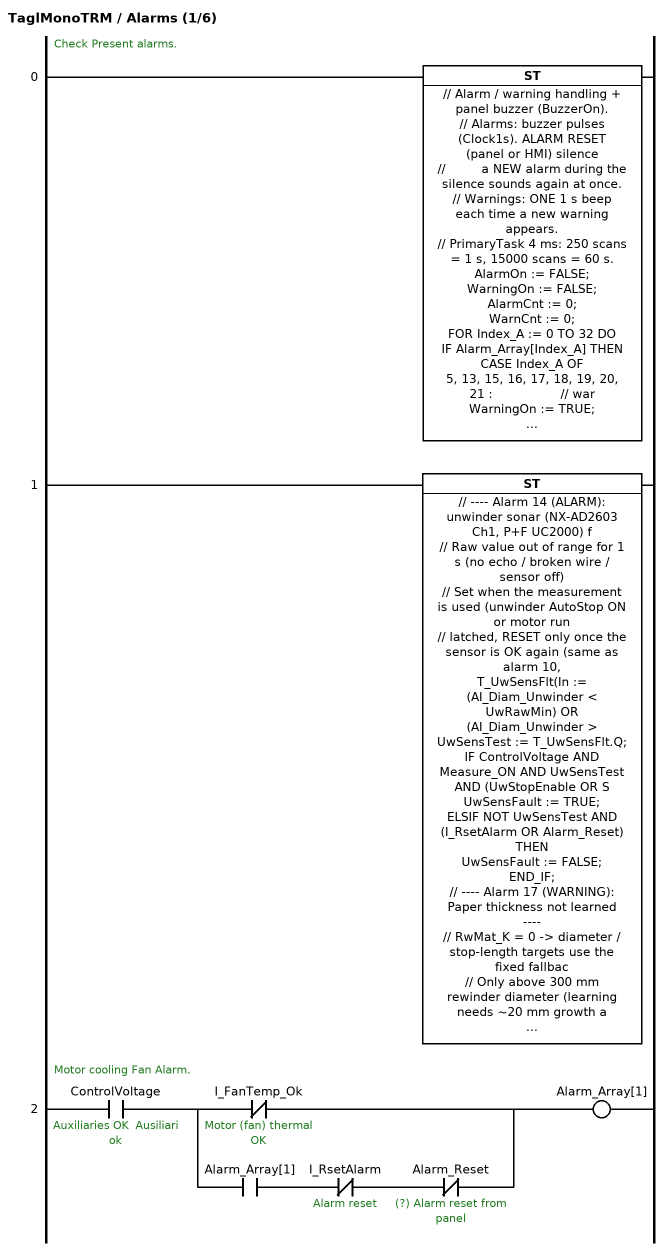
(* Rung 0: Check Present alarms. *)
// Alarm / warning handling + panel buzzer (BuzzerOn).
// Alarms: buzzer pulses (Clock1s). ALARM RESET (panel or HMI) silences it 1 min;
//         a NEW alarm during the silence sounds again at once.
// Warnings: ONE 1 s beep each time a new warning appears.
// PrimaryTask 4 ms: 250 scans = 1 s, 15000 scans = 60 s.

AlarmOn := FALSE;
WarningOn := FALSE;
AlarmCnt := 0;
WarnCnt := 0;

FOR Index_A := 0 TO 32 DO
	
    IF Alarm_Array[Index_A] THEN
        CASE Index_A OF
            5, 13, 15, 16, 17, 18, 19, 20, 21 :                 // warnings
                WarningOn := TRUE;
                WarnCnt := WarnCnt + 1;
        ELSE                          // alarms
            AlarmOn := TRUE;
            AlarmCnt := AlarmCnt + 1;
        END_CASE;
    END_IF;
END_FOR;

// ALARM RESET button (panel I_RsetAlarm or HMI Alarm_Reset): silence 1 min

RstEdge := (I_RsetAlarm OR Alarm_Reset) AND NOT RstMem;
RstMem := I_RsetAlarm OR Alarm_Reset;

IF RstEdge AND AlarmOn THEN
    SilenceTicks := 15000;
END_IF;

IF (AlarmCnt > AlarmCntMem) OR NOT AlarmOn THEN
    SilenceTicks := 0;                              // new alarm / no alarm: not silenced
END_IF;

IF SilenceTicks > 0 THEN
    SilenceTicks := SilenceTicks - 1;
END_IF;

// New warning: one 1 s beep

IF WarnCnt > WarnCntMem THEN
    WarnBeepTicks := 250;
END_IF;

IF WarnBeepTicks > 0 THEN
    WarnBeepTicks := WarnBeepTicks - 1;
END_IF;

AlarmCntMem := AlarmCnt;
WarnCntMem := WarnCnt;

AlarmSilenced := AlarmOn AND (SilenceTicks > 0);

BuzzerOn := ControlVoltage
            AND ((AlarmOn AND NOT AlarmSilenced AND Clock1s) OR (WarnBeepTicks > 0));
(* Rung 1 *)
// ---- Alarm 14 (ALARM): unwinder sonar (NX-AD2603 Ch1, P+F UC2000) fault ----
// Raw value out of range for 1 s (no echo / broken wire / sensor off).
// Set when the measurement is used (unwinder AutoStop ON or motor running),
// latched, RESET only once the sensor is OK again (same as alarm 10, DT35).

T_UwSensFlt(In := (AI_Diam_Unwinder < UwRawMin) OR (AI_Diam_Unwinder > UwRawMax), PT := T#1s);
UwSensTest := T_UwSensFlt.Q;

IF ControlVoltage AND Measure_ON AND UwSensTest AND (UwStopEnable OR StartMotor_Cmd) THEN
    UwSensFault := TRUE;
ELSIF NOT UwSensTest AND (I_RsetAlarm OR Alarm_Reset) THEN
    UwSensFault := FALSE;
END_IF;

// ---- Alarm 17 (WARNING): Paper thickness not learned ----
// RwMat_K = 0 -> diameter / stop-length targets use the fixed fallback.
// Only above 300 mm rewinder diameter (learning needs ~20 mm growth after NEW PAPER),
// so it does not beep at every new roll. Not latched.

Thickness_Fault := ControlVoltage AND StartMotor_Cmd 
                   AND (RwMat_K <= 0.0) AND (RwDiam > 300.0);
(* Rung 2: Motor cooling Fan Alarm. *)
Alarm_Array[1] := ControlVoltage AND (NOT I_FanTemp_Ok OR (Alarm_Array[1] AND NOT I_RsetAlarm AND NOT Alarm_Reset));

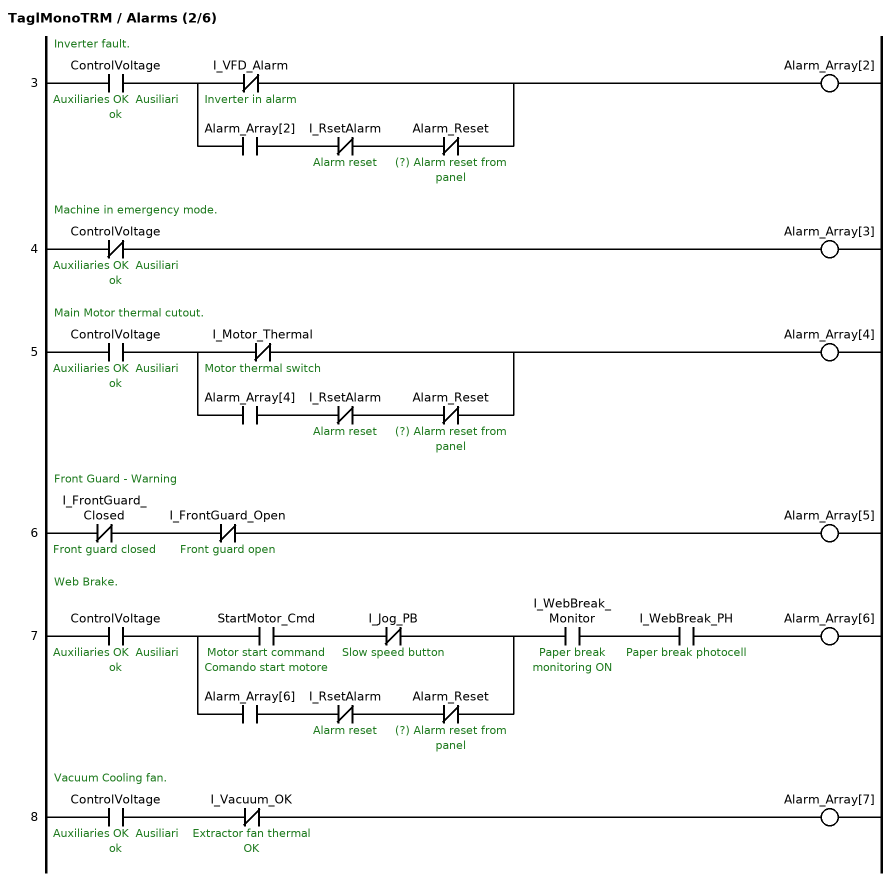
(* Rung 3: Inverter fault. *)
Alarm_Array[2] := ControlVoltage AND (NOT I_VFD_Alarm OR (Alarm_Array[2] AND NOT I_RsetAlarm AND NOT Alarm_Reset));
(* Rung 4: Machine in emergency mode. *)
Alarm_Array[3] := NOT ControlVoltage;
(* Rung 5: Main Motor thermal cutout. *)
Alarm_Array[4] := ControlVoltage AND (NOT I_Motor_Thermal OR (Alarm_Array[4] AND NOT I_RsetAlarm AND NOT Alarm_Reset));
(* Rung 6: Front Guard - Warning *)
Alarm_Array[5] := NOT I_FrontGuard_Closed AND NOT I_FrontGuard_Open;
(* Rung 7: Web Brake. *)
Alarm_Array[6] := ControlVoltage AND ((StartMotor_Cmd AND NOT I_Jog_PB) OR (Alarm_Array[6] AND NOT I_RsetAlarm AND NOT Alarm_Reset)) AND I_WebBreak_Monitor AND I_WebBreak_PH;
(* Rung 8: Vacuum Cooling fan. *)
Alarm_Array[7] := ControlVoltage AND NOT I_Vacuum_OK;

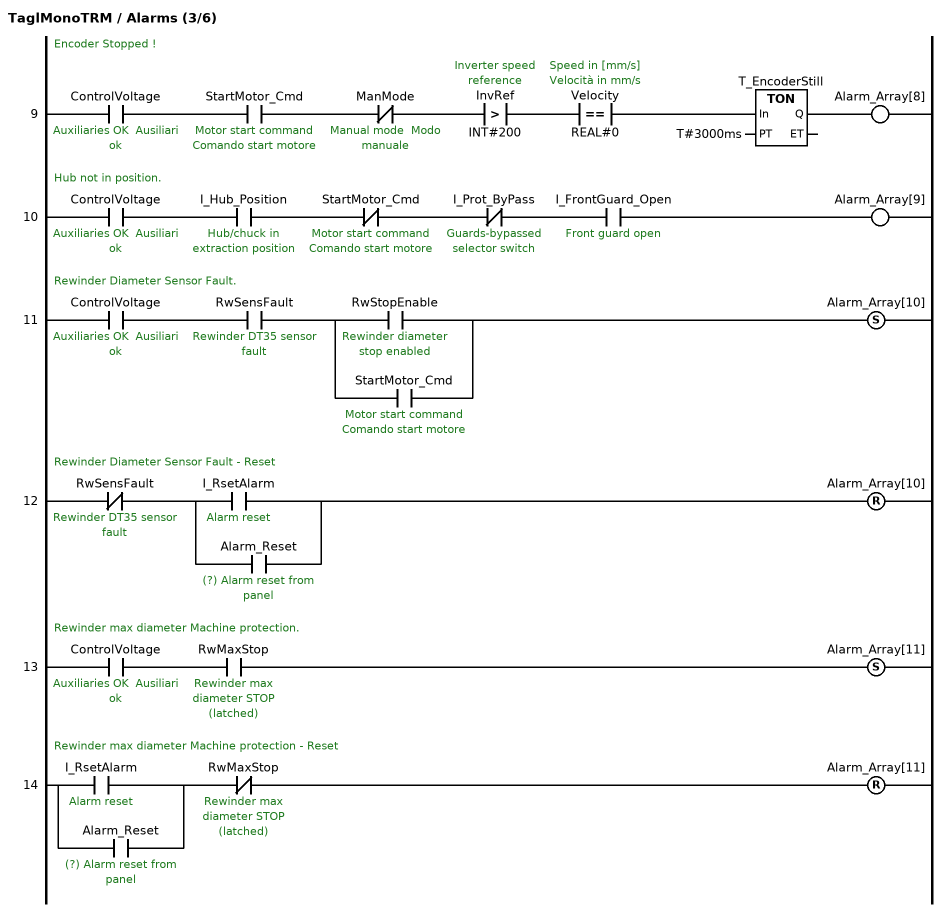
(* Rung 9: Encoder Stopped ! *)
T_EncoderStill(In := ControlVoltage AND StartMotor_Cmd AND NOT ManMode AND (InvRef > INT#200) AND (Velocity = REAL#0), PT := T#3000ms);
Alarm_Array[8] := T_EncoderStill.Q;
(* Rung 10: Hub not in position. *)
Alarm_Array[9] := ControlVoltage AND I_Hub_Position AND NOT StartMotor_Cmd AND NOT I_Prot_ByPass AND I_FrontGuard_Open;
(* Rung 11: Rewinder Diameter Sensor Fault. *)
IF ControlVoltage AND RwSensFault AND (RwStopEnable OR StartMotor_Cmd) THEN
    Alarm_Array[10] := TRUE;
END_IF;
(* Rung 12: Rewinder Diameter Sensor Fault - Reset *)
IF NOT RwSensFault AND (I_RsetAlarm OR Alarm_Reset) THEN Alarm_Array[10] := FALSE; END_IF;
(* Rung 13: Rewinder max diameter Machine protection. *)
IF ControlVoltage AND RwMaxStop THEN Alarm_Array[11] := TRUE; END_IF;
(* Rung 14: Rewinder max diameter Machine protection - Reset *)
IF (I_RsetAlarm OR Alarm_Reset) AND NOT RwMaxStop THEN Alarm_Array[11] := FALSE; END_IF;

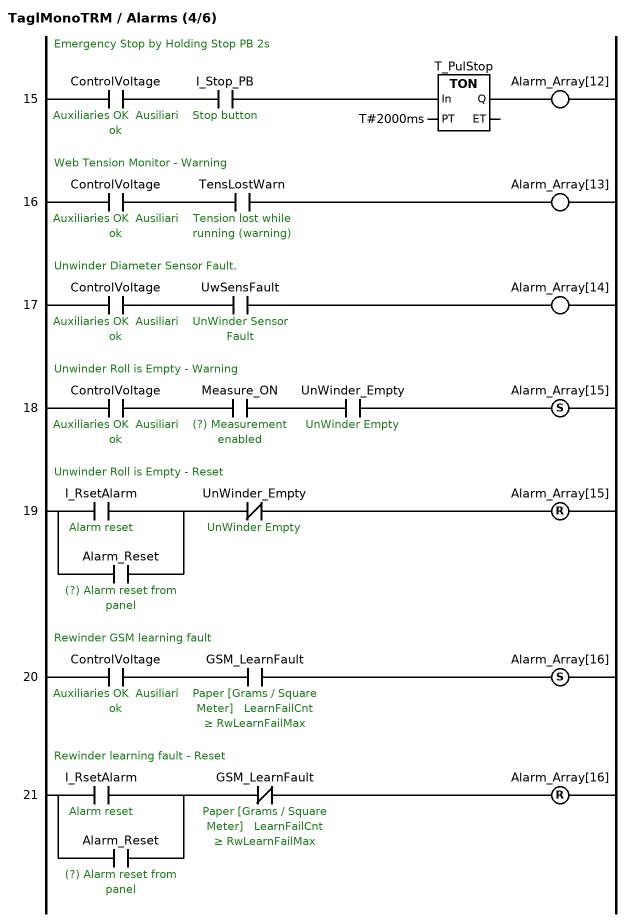
(* Rung 15: Emergency Stop by Holding Stop PB 2s *)
T_PulStop(In := ControlVoltage AND I_Stop_PB, PT := T#2000ms);
Alarm_Array[12] := T_PulStop.Q;
(* Rung 16: Web Tension Monitor - Warning *)
Alarm_Array[13] := ControlVoltage AND TensLostWarn;
(* Rung 17: Unwinder Diameter Sensor Fault. *)
Alarm_Array[14] := ControlVoltage AND UwSensFault;
(* Rung 18: Unwinder Roll is Empty - Warning *)
IF ControlVoltage AND Measure_ON AND UnWinder_Empty THEN Alarm_Array[15] := TRUE; END_IF;
(* Rung 19: Unwinder Roll is Empty - Reset *)
IF (I_RsetAlarm OR Alarm_Reset) AND NOT UnWinder_Empty THEN Alarm_Array[15] := FALSE; END_IF;
(* Rung 20: Rewinder GSM learning fault *)
IF ControlVoltage AND GSM_LearnFault THEN Alarm_Array[16] := TRUE; END_IF;
(* Rung 21: Rewinder learning fault - Reset *)
IF (I_RsetAlarm OR Alarm_Reset) AND NOT GSM_LearnFault THEN Alarm_Array[16] := FALSE; END_IF;

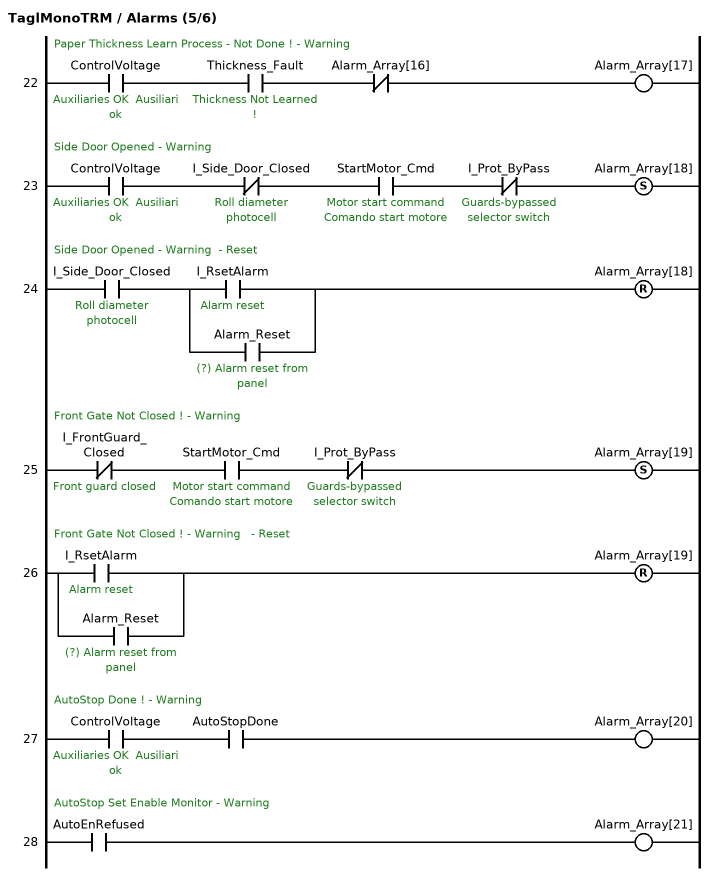
(* Rung 22: Paper Thickness Learn Process - Not Done ! - Warning *)
Alarm_Array[17] := ControlVoltage AND Thickness_Fault AND NOT Alarm_Array[16];
(* Rung 23: Side Door Opened - Warning *)
IF ControlVoltage AND NOT I_Side_Door_Closed AND StartMotor_Cmd AND NOT I_Prot_ByPass THEN
    Alarm_Array[18] := TRUE;
END_IF;
(* Rung 24: Side Door Opened - Warning  - Reset *)
IF I_Side_Door_Closed AND (I_RsetAlarm OR Alarm_Reset) THEN Alarm_Array[18] := FALSE; END_IF;
(* Rung 25: Front Gate Not Closed ! - Warning *)
IF NOT I_FrontGuard_Closed AND StartMotor_Cmd AND NOT I_Prot_ByPass THEN Alarm_Array[19] := TRUE; END_IF;
(* Rung 26: Front Gate Not Closed ! - Warning   - Reset *)
IF I_RsetAlarm OR Alarm_Reset THEN Alarm_Array[19] := FALSE; END_IF;
(* Rung 27: AutoStop Done ! - Warning *)
Alarm_Array[20] := ControlVoltage AND AutoStopDone;
(* Rung 28: AutoStop Set Enable Monitor - Warning *)
Alarm_Array[21] := AutoEnRefused;

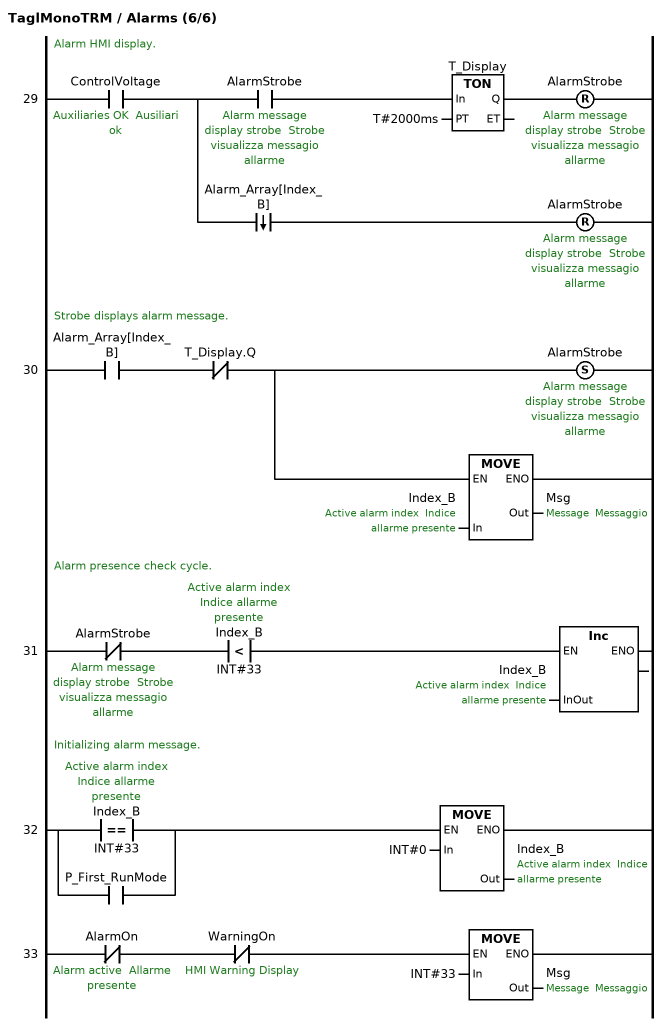
(* Rung 29: Alarm HMI display. *)
T_Display(In := ControlVoltage AND AlarmStrobe, PT := T#2000ms);
IF T_Display.Q THEN AlarmStrobe := FALSE; END_IF;
_e14(CLK := Alarm_Array[Index_B]);
IF ControlVoltage AND _e14.Q THEN AlarmStrobe := FALSE; END_IF;
(* Rung 30: Strobe displays alarm message. *)
IF Alarm_Array[Index_B] AND NOT T_Display.Q THEN
    AlarmStrobe := TRUE;
    Msg := Index_B;
END_IF;
(* Rung 31: Alarm presence check cycle. *)
IF NOT AlarmStrobe AND (Index_B < INT#33) THEN Inc(InOut := Index_B); END_IF;
(* Rung 32: Initializing alarm message. *)
IF (Index_B = INT#33) OR P_First_RunMode THEN Index_B := INT#0; END_IF;
(* Rung 33 *)
IF NOT AlarmOn AND NOT WarningOn THEN Msg := INT#33; END_IF;

(* Section Output_Manager: ladder, written here as Structured Text *)

